(* IEC 61131-3 sources: daoli-st-library/DL_Device (part 8) *)

(* ---- FC_DL_BatteryBackupTimeCalc.st ---- *)
(*
 * FC_DL_BatteryBackupTimeCalc | C2 | DL_Device
 * 功能：电池组恒功率放电后备时间（含寿命末期与放电效率修正）       单位：容量 [Ah]、电压 [V]、功率 [kW]、时间 [min]、修正系数 [1]
 * 工况边界：恒功率简化模型（不含 Peukert 效应与温度修正，温度影响由 rDerate 吸收）；负载功率须 >0（入分母），容量、电压须 >0，两修正系数须在 (0,1]；电池组按串联单体电压和计算
 * 代数值回代：C=200 Ah、V=480 V、P=100 kW、derate=0.85、eol=0.8 → 200×480×0.85×0.8=65280 Wh；65280/100000=0.6528 h=39.17 min（spec 记 39.2 min，一致）
 * 开源溯源：clean-room 自研，未复制任何第三方代码（无外部来源）
 *)
FUNCTION FC_DL_BatteryBackupTimeCalc : BOOL
VAR_INPUT
    rCapacityAh : REAL := 200.0;     // 电池组额定容量 | battery string rated capacity [Ah]
    rStringV    : REAL := 480.0;     // 电池组标称电压 | battery string nominal voltage [V]
    rLoadKw     : REAL := 100.0;     // 放电负载功率 | discharge load power [kW]
    rDerate     : REAL := 0.85;      // 放电效率与温度综合修正 | combined discharge efficiency and temperature derating [1]
    rEolFactor  : REAL := 0.8;       // 寿命末期容量保持率 | end of life capacity retention [1]
END_VAR
VAR_OUTPUT
    rBackupMin : REAL;               // 后备时间 | backup time [min]
    rEnergyWh  : REAL;               // 可用能量 | usable energy [Wh]
    xValid     : BOOL;               // 输出有效 | outputs valid
END_VAR
VAR
    xFinC   : BOOL;                  // 容量有限性 | capacity is finite
    xFinV   : BOOL;                  // 电压有限性 | voltage is finite
    xFinP   : BOOL;                  // 功率有限性 | load power is finite
    xFinDr  : BOOL;                  // 效率修正有限性 | derating factor is finite
    xFinEol : BOOL;                  // 寿命修正有限性 | end of life factor is finite
    rPW     : REAL;                  // 负载功率（W）| load power in watts [W]
END_VAR
VAR CONSTANT
    DL_BBT_MIN_PER_HOUR : REAL := 60.0;    // 小时转分系数 | hours to minutes factor [min/h]
    DL_BBT_W_PER_KW     : REAL := 1000.0;  // 千瓦转瓦系数 | kilowatts to watts factor [W/kW]
    DL_BBT_P_MIN        : REAL := 1.0E-9;  // 负载功率下限（防零除）| load power lower bound [W]
END_VAR

// 段1｜非有限闸（R19）
xFinC := (rCapacityAh = rCapacityAh) AND ((rCapacityAh - rCapacityAh) = 0.0);
xFinV := (rStringV = rStringV) AND ((rStringV - rStringV) = 0.0);
xFinP := (rLoadKw = rLoadKw) AND ((rLoadKw - rLoadKw) = 0.0);
xFinDr := (rDerate = rDerate) AND ((rDerate - rDerate) = 0.0);
xFinEol := (rEolFactor = rEolFactor) AND ((rEolFactor - rEolFactor) = 0.0);
IF (NOT xFinC) OR (NOT xFinV) OR (NOT xFinP) OR (NOT xFinDr) OR (NOT xFinEol) THEN
    rBackupMin := 0.0;               // 安全值：后备时间 0 | safe value, zero backup time
    rEnergyWh := 0.0;
    xValid := FALSE;
    FC_DL_BatteryBackupTimeCalc := FALSE;
    RETURN;
END_IF

// 段2｜域闸：容量/电压/功率须为正，两修正系数须在 (0,1]
IF (rCapacityAh <= 0.0) OR (rStringV <= 0.0) OR (rLoadKw <= 0.0)
   OR (rDerate <= 0.0) OR (rDerate > 1.0) OR (rEolFactor <= 0.0) OR (rEolFactor > 1.0) THEN
    rBackupMin := 0.0;
    rEnergyWh := 0.0;
    xValid := FALSE;
    FC_DL_BatteryBackupTimeCalc := FALSE;
    RETURN;
END_IF

// 段3｜算法：可用能量 Wh 与后备时间 min
rEnergyWh := rCapacityAh * rStringV * rDerate * rEolFactor;
rPW := rLoadKw * DL_BBT_W_PER_KW;
IF rPW > DL_BBT_P_MIN THEN
    rBackupMin := rEnergyWh / rPW * DL_BBT_MIN_PER_HOUR;
ELSE
    rBackupMin := 0.0;               // 理论不可达（段2已排除），防御性兜底 | unreachable defence
END_IF

// 段4｜出口
xValid := TRUE;
FC_DL_BatteryBackupTimeCalc := TRUE;
END_FUNCTION

(* ---- FC_DL_BoothFilterLifeCalc.st ---- *)
(*
  Name: FC_DL_BoothFilterLifeCalc
  Category: DL_Device
  Version: 1.0.0
  Round: R89 / 2026-11-25
  开源溯源：clean-room 自研（族 涂装喷涂线，ST 开源生态实测 0 命中，无外部代码引入）
  功能：过滤棉剩余寿命：按压差累积法算寿命消耗百分比，并按当前压差增长率外推剩余运行小时。
  边界条件：① 四入参全部过非有限闸，任一非有限返回哨兵 -1；
            ② 新棉压差必须 > 0 且报废压差必须高于新棉压差（否则分母 ΔP 塌零，返回哨兵 -1）；
            ③ 已用压差 Δp − Δp_new 为除子，外推前显式判零：低于 DL_EPS 时剩余小时按满寿命处理；
            ④ 寿命百分比钳 0~100 %（量值饱和）；报警门限 90 %，超报废压差即 100 % 并报警。
  量纲自证：(ΔP − ΔP_new)/(ΔP_end − ΔP_new) 无量纲；h × 无量纲 = h。
*)
FUNCTION FC_DL_BoothFilterLifeCalc : REAL
VAR_INPUT
    fDpPa : REAL;           (* 当前滤棉压差 [Pa] Current filter pressure drop [Pa] *)
    fDpNewPa : REAL;        (* 新棉压差（洁净基线） [Pa] Clean filter pressure drop [Pa] *)
    fDpEndPa : REAL;        (* 报废压差 [Pa] End-of-life pressure drop [Pa] *)
    fRunHours : REAL;       (* 滤棉已运行小时 [h] Filter accumulated run hours [h] *)
END_VAR
VAR_OUTPUT
    fLifeUsedPct : REAL;    (* 寿命消耗百分比 [%] Life used [%] *)
    fRemainHours : REAL;    (* 剩余可用小时（外推） [h] Remaining hours, extrapolated [h] *)
    xReplaceAlarm : BOOL;   (* 更换报警（寿命 ≥ 90 %） [-] Replace alarm *)
    xValid : BOOL;          (* 计算有效性标志 [-] Calculation valid flag *)
END_VAR
VAR CONSTANT
    DL_EPS : REAL := 1.0E-9;        (* 除零判定容差 [-] Divide-by-zero tolerance *)
    DL_PCT : REAL := 100.0;         (* 百分数基准 [%] Percent base *)
    DL_ALARM_PCT : REAL := 90.0;    (* 更换报警门限 [%] Replace alarm threshold [%] *)
    DL_P_NEW_MAX : REAL := 500.0;   (* 新棉压差上限 [Pa] Clean pressure ceiling [Pa] *)
    DL_P_END_MIN : REAL := 100.0;   (* 报废压差下限 [Pa] End pressure floor [Pa] *)
    DL_P_END_MAX : REAL := 5000.0;  (* 报废压差上限 [Pa] End pressure ceiling [Pa] *)
    DL_H_MAX : REAL := 100000.0;    (* 运行小时上限 [h] Run hours ceiling [h] *)
END_VAR
VAR
    fSpanPa : REAL;     (* 全寿命压差跨度 [Pa] Full-life pressure span [Pa] *)
    fUsedPa : REAL;     (* 已消耗压差 [Pa] Consumed pressure drop [Pa] *)
    fPct : REAL;        (* 寿命消耗中间量 [%] Life used scratch [%] *)
END_VAR
(* 出口预置：四出口统一预置（R256） *)
fLifeUsedPct := 0.0; fRemainHours := 0.0; xReplaceAlarm := FALSE; xValid := FALSE;
(* 非有限闸：NaN 自反判 + Inf 差值自减判，四入参全枚举 *)
IF (fDpPa <> fDpPa) OR ((fDpPa - fDpPa) <> 0.0)
   OR (fDpNewPa <> fDpNewPa) OR ((fDpNewPa - fDpNewPa) <> 0.0)
   OR (fDpEndPa <> fDpEndPa) OR ((fDpEndPa - fDpEndPa) <> 0.0)
   OR (fRunHours <> fRunHours) OR ((fRunHours - fRunHours) <> 0.0) THEN
    FC_DL_BoothFilterLifeCalc := -1.0;      (* 哨兵 -1：入参非有限 / Sentinel -1, non-finite input *)
    RETURN;
END_IF
(* 组态域闸：压差三点与运行小时定域，报废压差须高于新棉压差 *)
IF (fDpNewPa < DL_EPS) OR (fDpNewPa > DL_P_NEW_MAX)
   OR (fDpEndPa < DL_P_END_MIN) OR (fDpEndPa > DL_P_END_MAX)
   OR ((fDpEndPa - fDpNewPa) <= DL_EPS)
   OR (fDpPa < 0.0) OR (fDpPa > (fDpEndPa * 1.5))
   OR (fRunHours < 0.0) OR (fRunHours > DL_H_MAX) THEN
    FC_DL_BoothFilterLifeCalc := -1.0;      (* 哨兵 -1：组态非法 / Sentinel -1, bad configuration *)
    RETURN;
END_IF
(* 全寿命压差跨度已过正性闸，绝无零除 *)
fSpanPa := fDpEndPa - fDpNewPa;
(* 已消耗压差：低于新棉基线按 0 处理（新棉初期压差抖动不产生负寿命） *)
fUsedPa := fDpPa - fDpNewPa;
IF fUsedPa < 0.0 THEN
    fUsedPa := 0.0;
END_IF
(* 寿命消耗百分比 *)
fPct := (fUsedPa / fSpanPa) * DL_PCT;
IF fPct > DL_PCT THEN
    fPct := DL_PCT;                         (* 量值饱和：超报废压差即 100 % / Saturation at 100 % *)
END_IF
fLifeUsedPct := fPct;
(* 剩余小时外推：h × (剩余压差/已耗压差)；已耗压差塌零时按满寿命 + 无穷处置为 0 剩余待定 *)
IF fUsedPa <= DL_EPS THEN
    fRemainHours := DL_H_MAX;               (* 近乎新棉：剩余小时按可表上限 / Effectively new filter *)
ELSE
    fRemainHours := fRunHours * ((fSpanPa - fUsedPa) / fUsedPa);
    IF fRemainHours < 0.0 THEN
        fRemainHours := 0.0;                (* 已超报废压差：剩余 0 h / Past end of life *)
    END_IF
END_IF
xReplaceAlarm := fLifeUsedPct >= DL_ALARM_PCT;
xValid := TRUE;                             (* 链路有效 / Chain valid *)
FC_DL_BoothFilterLifeCalc := fLifeUsedPct;
END_FUNCTION

(* ---- FC_DL_BrgThermalDriftRate.st ---- *)
(*
  道莅工业代码库 / Daoli Industrial ST Library
  组件: FC_DL_BrgThermalDriftRate
  分类: DL_Device
  开源溯源: 无（clean-room 工程公式自研；参考公开工艺计算公式，未复制任何受版权保护代码）
  许可证: 本项目自有 (MIT)
  功能: 轴承温升速率计算、相对环境温升与温升过快判定
*)
FUNCTION FC_DL_BrgThermalDriftRate : BOOL
VAR_INPUT
    rTempNow : REAL; // 本次轴承温度 [°C] / current bearing temperature
    rTempPrev : REAL; // 上次轴承温度 [°C] / previous bearing temperature
    rDtMin : REAL; // 采样间隔 [min] / sampling interval in minutes
    rAmbC : REAL; // 环境温度 [°C] / ambient temperature
    rAlarmRisePerMin : REAL; // 温升速率报警门槛 [°C/min] / rise rate alarm threshold
END_VAR
VAR_OUTPUT
    rRisePerMin : REAL; // 温升速率 [°C/min] / temperature rise rate
    rOverAmbC : REAL; // 相对环境温升 [°C] / temperature rise above ambient
    bValid : BOOL; // 结果有效位 [-] / result valid flag
    bFastRise : BOOL; // 温升过快标志 [-] / fast rise flag
    iErrCode : INT; // 事件码 0=正常 1=采样间隔非法 2=结果非有限 / event code
END_VAR
VAR CONSTANT
    rAbsZero : REAL := -273.15; // 绝对零度 [°C] / absolute zero in Celsius
END_VAR
VAR
    rRiseRaw : REAL; // 未校验温升速率 [°C/min] / unchecked rise rate
END_VAR

    // —— 段 0：全路径预清 —— //
    rRiseRaw := 0.0;
    rRisePerMin := 0.0;
    rOverAmbC := 0.0;
    bValid := FALSE;
    bFastRise := FALSE;
    iErrCode := 0;
    FC_DL_BrgThermalDriftRate := FALSE;
    // —— 段 1：分母闸（采样间隔必须为正） —— //
    IF rDtMin <= 0.0 THEN
        iErrCode := 1; // 采样间隔非法，速率无定义 / invalid interval, rate undefined
        RETURN;
    END_IF;
    // —— 段 2：量纲链 (°C - °C)/(min) = °C/min —— //
    rRiseRaw := (rTempNow - rTempPrev) / rDtMin; // 温升速率 [°C/min] / rise rate
    IF ABS(rRiseRaw) > 1.0E15 THEN
        iErrCode := 2; // 结果非有限，强制归零 / non-finite result, forced to zero
        RETURN;
    END_IF;
    rRisePerMin := rRiseRaw;
    // —— 段 3：相对环境温升（量纲 °C - °C = °C） —— //
    IF rTempNow <= rAbsZero THEN
        iErrCode := 2; // 温度低于绝对零度，物理不可能 / temperature below absolute zero
        RETURN;
    END_IF;
    rOverAmbC := rTempNow - rAmbC; // 相对环境温升 [°C] / rise above ambient
    // —— 段 4：温升过快判定（门槛为负时按绝对值口径比对） —— //
    IF rAlarmRisePerMin > 0.0 THEN
        bFastRise := rRisePerMin > rAlarmRisePerMin; // 常规比对 / normal comparison
    ELSE
        bFastRise := rRisePerMin > ABS(rAlarmRisePerMin); // 门槛配置异常时退化为绝对值口径 / fallback on bad threshold
    END_IF;
    bValid := TRUE;
    FC_DL_BrgThermalDriftRate := TRUE;
END_FUNCTION

(* ---- FC_DL_BushingDwellFlowCalc.st ---- *)
// FC_DL_BushingDwellFlowCalc v1.0.0
// 开源溯源：clean-room 自研（族 DL_Device，ST 生态实测 0 命中，无外部代码引入）
(*
  功能: 漏孔玻璃液质量流量（Hagen-Poiseuille 圆管层流）：r = d/2/1000，L = len/1000，
        Q = π·Δp·r⁴/(8·μ·L) [m³/s]，单孔 = Q·ρ·3.6e6 [g/h]，总流量 = 单孔·孔数/1000 [kg/h]。
  邻件/码位: 与 FC_DL_FiberDiameterFromDrawRateCalc 直接串联（本件出单孔流量）；
             16#0002_9222 = 非有限、黏度/孔径/孔长/密度非正或孔数 < 1 拒收。
*)
FUNCTION FC_DL_BushingDwellFlowCalc : REAL
VAR_INPUT
    fDeltaP    : REAL := 5000.0;    // 漏板上下压差 [Pa]，域 > 0 / Pressure differential [Pa]
    fHoleDia   : REAL := 1.6;       // 漏孔直径 [mm]，域 > 0 / Orifice diameter [mm]
    fDwellLen  : REAL := 4.0;       // 漏孔长度 [mm]，域 > 0 / Orifice length [mm]
    fViscosity : REAL := 500.0;     // 玻璃液黏度 [Pa·s]，域 > 0 / Glass viscosity [Pa s]
    iHoleCount : INT := 800;        // 漏孔数，域 >= 1 [个] / Orifice count
    fDensity   : REAL := 2500.0;    // 玻璃液密度 [kg/m³]，域 > 0 / Glass density [kg/m^3]
END_VAR
VAR_OUTPUT
    fFlowPerHole : REAL;            // 单孔质量流量 [g/h] / Mass flow per orifice [g/h]
    fFlowTotal   : REAL;            // 总质量流量 [kg/h] / Total mass flow [kg/h]
    bValid       : BOOL;            // 结果有效回执 [-] / Result validity receipt
    uErrorId     : UDINT;           // 事件码，0 = 无事件 / Event code
END_VAR
VAR
    fRadius  : REAL := 0.0;         // 漏孔半径 [m] / Orifice radius [m]
    fLenM    : REAL := 0.0;         // 漏孔长度 [m] / Orifice length [m]
    fVolFlow : REAL := 0.0;         // 单孔体积流量 [m³/s] / Volumetric flow [m^3/s]
END_VAR
// 段 0：全路径出口安全缺省 / Safe defaults on all outlets
fFlowPerHole := 0.0;                // 单孔流量缺省零 / Per-orifice default zero
fFlowTotal := 0.0;                  // 总流量缺省零 / Total flow default zero
bValid := FALSE;                    // 有效回执预清 / Validity preset clear
uErrorId := 16#0000;                // 事件码预清 / Event code preset clear
FC_DL_BushingDwellFlowCalc := 0.0;  // 返回值缺省零（镜像单孔流量）/ Return default zero
// 段 1：非有限闸（五实数入参；整数入参天然有限）/ Non-finite gate on real inputs
IF (fDeltaP <> fDeltaP) OR (fHoleDia <> fHoleDia) OR (fDwellLen <> fDwellLen)
   OR (fViscosity <> fViscosity) OR (fDensity <> fDensity)
   OR (ABS(fDeltaP) >= 3.0E38) OR (ABS(fHoleDia) >= 3.0E38) OR (ABS(fDwellLen) >= 3.0E38)
   OR (ABS(fViscosity) >= 3.0E38) OR (ABS(fDensity) >= 3.0E38) THEN
    uErrorId := 16#0002_9222;   // 入参非有限拒收 / Non-finite input reject
    RETURN;
END_IF
// 段 2：域闸（黏度/孔径/孔长/密度为正防除零 + 孔数下限，R4）/ Domain gate
IF (fViscosity <= 1.0E-6) OR (fHoleDia <= 1.0E-6) OR (fDwellLen <= 1.0E-6) OR (fDensity <= 1.0E-6) THEN
    uErrorId := 16#0002_9222;   // 黏度、孔径、孔长或密度非正 / Non-positive physical input
    RETURN;
END_IF
IF iHoleCount < 1 THEN
    uErrorId := 16#0002_9222;   // 孔数不足 1 / Orifice count below one
    RETURN;
END_IF
// 段 3：主计算（半径/长度换算 → 体积流量 → 质量流量）/ Main computation
fRadius := fHoleDia / 2.0 / 1000.0;                             // 半径 [m] / Radius in metres
fLenM := fDwellLen / 1000.0;                                    // 孔长 [m] / Length in metres
fVolFlow := 3.14159265358979 * fDeltaP * fRadius * fRadius * fRadius * fRadius
          / (8.0 * fViscosity * fLenM);                         // Q = πΔp r⁴/(8μL) / Poiseuille flow
fFlowPerHole := fVolFlow * fDensity * 3600.0 * 1000.0;          // 单孔 [g/h] / Per-orifice mass flow
fFlowTotal := fFlowPerHole * INT_TO_REAL(iHoleCount) / 1000.0;  // 总流量 [kg/h] / Total mass flow
// 段 4：出口闸（双输出非有限复核 + 非负复核）/ Outlet gate
IF (fFlowPerHole <> fFlowPerHole) OR (fFlowTotal <> fFlowTotal)
   OR (ABS(fFlowPerHole) >= 3.0E38) OR (ABS(fFlowTotal) >= 3.0E38)
   OR (fFlowPerHole < 0.0) OR (fFlowTotal < 0.0) THEN
    fFlowPerHole := 0.0;        // 复核失败回缺省 / Fallback on recheck failure
    fFlowTotal := 0.0;          // 复核失败回缺省 / Fallback on recheck failure
    uErrorId := 16#0002_9222;   // 出口复核拒收 / Output recheck reject
    RETURN;
END_IF
bValid := TRUE;                 // 有效回执 / Validity receipt
FC_DL_BushingDwellFlowCalc := fFlowPerHole;     // 返回值镜像单孔流量 / Return mirrors flow
END_FUNCTION

(* ---- FC_DL_BushingPowerBalanceCalc.st ---- *)
// FC_DL_BushingPowerBalanceCalc v1.0.0
// 开源溯源：clean-room 自研（族 DL_Device，ST 生态实测 0 命中，无外部代码引入）
(*
  功能: 漏板电热功率平衡：输入功率 = I²·R [W]→[kW]（mΩ 除 1000 转 Ω，W 除 1000 转 kW），
        对流 = 12·A·ΔT/1000 [kW]（12 为自然对流综合换热系数 W/(m²·K)），
        辐射 = εσ·A·(T_K⁴ − Ta_K⁴)/1000 [kW]（ε = 0.85，σ = 5.67e-8），
        热效率 = 1 − (对流 + 辐射)/输入功率。
  邻件/码位: 与 FC_DL_BushingTempZoneCalc 为热平衡两侧（温度设定 vs 实际电功率与散热）；
             16#0002_9227 = 非有限、电阻/面积非正、温度不高于绝对零度、输入功率近零或效率出物理域。
*)
FUNCTION FC_DL_BushingPowerBalanceCalc : REAL
VAR_INPUT
    fCurrent     : REAL := 300.0;   // 漏板电流 [A]，域 > 0 / Bushing current [A]
    fResistance  : REAL := 30.0;    // 漏板电阻 [mΩ]，域 > 0 / Bushing resistance [mOhm]
    fSurfaceArea : REAL := 0.5;     // 漏板表面积 [m²]，域 > 0 / Surface area [m^2]
    fTemp        : REAL := 1200.0;  // 漏板温度 [°C] / Bushing temperature [degC]
    fAmbient     : REAL := 30.0;    // 环境温度 [°C] / Ambient temperature [degC]
END_VAR
VAR_OUTPUT
    fPowerIn    : REAL;             // 输入电功率 [kW] / Electrical input power [kW]
    fLossConv   : REAL;             // 对流散热 [kW] / Convective loss [kW]
    fLossRad    : REAL;             // 辐射散热 [kW] / Radiative loss [kW]
    fEfficiency : REAL;             // 热效率 [-] / Thermal efficiency
    bValid      : BOOL;             // 结果有效回执 [-] / Result validity receipt
    uErrorId    : UDINT;            // 事件码，0 = 无事件 / Event code
END_VAR
VAR
    fTK  : REAL := 0.0;             // 板绝对温度 [K] / Bushing absolute temperature [K]
    fTaK : REAL := 0.0;             // 环境绝对温度 [K] / Ambient absolute temperature [K]
END_VAR
// 段 0：全路径出口安全缺省 / Safe defaults on all outlets
fPowerIn := 0.0;                    // 输入功率缺省零 / Input power default zero
fLossConv := 0.0;                   // 对流散热缺省零 / Convective loss default zero
fLossRad := 0.0;                    // 辐射散热缺省零 / Radiative loss default zero
fEfficiency := 0.0;                 // 热效率缺省零 / Efficiency default zero
bValid := FALSE;                    // 有效回执预清 / Validity preset clear
uErrorId := 16#0000;                // 事件码预清 / Event code preset clear
FC_DL_BushingPowerBalanceCalc := 0.0;   // 返回值缺省零（镜像热效率）/ Return default zero
// 段 1：非有限闸（五入参全枚举）/ Non-finite gate over all inputs
IF (fCurrent <> fCurrent) OR (fResistance <> fResistance) OR (fSurfaceArea <> fSurfaceArea)
   OR (fTemp <> fTemp) OR (fAmbient <> fAmbient)
   OR (ABS(fCurrent) >= 3.0E38) OR (ABS(fResistance) >= 3.0E38) OR (ABS(fSurfaceArea) >= 3.0E38)
   OR (ABS(fTemp) >= 3.0E38) OR (ABS(fAmbient) >= 3.0E38) THEN
    uErrorId := 16#0002_9227;   // 入参非有限拒收 / Non-finite input reject
    RETURN;
END_IF
// 段 2：域闸（电阻/面积为正 + 温度高于绝对零度 + 输入功率近零，R4）/ Domain gate
IF (fResistance <= 1.0E-6) OR (fSurfaceArea <= 1.0E-6) THEN
    uErrorId := 16#0002_9227;   // 电阻或面积非正 / Non-positive resistance or area
    RETURN;
END_IF
IF (fTemp <= -273.15) OR (fAmbient <= -273.15) THEN
    uErrorId := 16#0002_9227;   // 温度不高于绝对零度，四次方无意义 / At or below absolute zero
    RETURN;
END_IF
fPowerIn := fCurrent * fCurrent * (fResistance / 1000.0) / 1000.0;      // I²R [kW] / Input power
IF fPowerIn <= 1.0E-6 THEN
    uErrorId := 16#0002_9227;   // 输入功率近零，效率不可解 / Input power too small
    RETURN;
END_IF
// 段 3：主计算（对流 + 辐射 + 效率）/ Main computation
fTK := fTemp + 273.15;                                          // 板绝对温度 [K] / Absolute temperature
fTaK := fAmbient + 273.15;                                      // 环境绝对温度 [K] / Ambient absolute temperature
fLossConv := 12.0 * fSurfaceArea * (fTemp - fAmbient) / 1000.0;  // 对流散热 [kW] / Convective loss
fLossRad := 5.67E-8 * 0.85 * fSurfaceArea * ((fTK * fTK * fTK * fTK) - (fTaK * fTaK * fTaK * fTaK)) / 1000.0;
fEfficiency := 1.0 - (fLossConv + fLossRad) / fPowerIn;         // 热效率 / Thermal efficiency
// 段 4：出口闸（四输出非有限复核 + 效率区间复核）/ Outlet gate
IF (fPowerIn <> fPowerIn) OR (fLossConv <> fLossConv) OR (fLossRad <> fLossRad)
   OR (fEfficiency <> fEfficiency)
   OR (ABS(fPowerIn) >= 3.0E38) OR (ABS(fLossConv) >= 3.0E38)
   OR (ABS(fLossRad) >= 3.0E38) OR (ABS(fEfficiency) >= 3.0E38) THEN
    fPowerIn := 0.0;            // 复核失败回缺省 / Fallback on recheck failure
    fLossConv := 0.0;           // 复核失败回缺省 / Fallback on recheck failure
    fLossRad := 0.0;            // 复核失败回缺省 / Fallback on recheck failure
    fEfficiency := 0.0;         // 复核失败回缺省 / Fallback on recheck failure
    uErrorId := 16#0002_9227;   // 出口非有限拒收 / Output non-finite reject
    RETURN;
END_IF
IF (fEfficiency > 1.0) OR (fEfficiency < -1.0) THEN
    uErrorId := 16#0002_9227;   // 信息级：效率出物理域 / Info: efficiency out of physical range
    RETURN;                     // bValid 保持 FALSE / Validity stays false
END_IF
bValid := TRUE;                 // 有效回执 / Validity receipt
FC_DL_BushingPowerBalanceCalc := fEfficiency;   // 返回值镜像热效率 / Return mirrors efficiency
END_FUNCTION

(* ---- FC_DL_BushingTempZoneCalc.st ---- *)
// FC_DL_BushingTempZoneCalc v1.0.0
// 开源溯源：clean-room 自研（族 DL_Device，ST 生态实测 0 命中，无外部代码引入）
(*
  功能: 漏板分区温度设定：偏移 = 梯度·(iZoneIndex − (iZoneCount−1)/2)，温度 = 基准 + 偏移；
        以区号相对中心对称取偏移，保证漏板横向温度对称分布。
  邻件/码位: 与 FC_DL_BushingDwellFlowCalc（温度→黏度→流量）上游衔接；
             16#0002_9221 = 非有限、区数非正、区号越界或温度出 1100~1350 °C 拒收。
*)
FUNCTION FC_DL_BushingTempZoneCalc : REAL
VAR_INPUT
    fBaseTemp  : REAL := 1250.0;    // 中心区设定温度 [°C] / Center zone setpoint [degC]
    fGradient  : REAL := 5.0;       // 区间梯度 [°C/区] / Per-zone gradient [degC/zone]
    iZoneIndex : INT := 0;          // 区号，0 起 [-] / Zone index, zero based
    iZoneCount : INT := 1;          // 总区数，域 > 0 [-] / Total zone count
END_VAR
VAR_OUTPUT
    fZoneTemp : REAL;               // 分区温度设定 [°C] / Zone temperature setpoint [degC]
    bValid    : BOOL;               // 结果有效回执 [-] / Result validity receipt
    uErrorId  : UDINT;              // 事件码，0 = 无事件 / Event code
END_VAR
VAR
    fCenter : REAL := 0.0;          // 中心区号（可为半整数）[-] / Center zone position
END_VAR
// 段 0：全路径出口安全缺省 / Safe defaults on all outlets
fZoneTemp := 0.0;               // 分区温度缺省零 / Zone temperature default zero
bValid := FALSE;                // 有效回执预清 / Validity preset clear
uErrorId := 16#0000;            // 事件码预清 / Event code preset clear
FC_DL_BushingTempZoneCalc := 0.0;       // 返回值缺省零（镜像分区温度）/ Return default zero
// 段 1：非有限闸（两实数入参；整数入参天然有限）/ Non-finite gate on real inputs
IF (fBaseTemp <> fBaseTemp) OR (fGradient <> fGradient)
   OR (ABS(fBaseTemp) >= 3.0E38) OR (ABS(fGradient) >= 3.0E38) THEN
    uErrorId := 16#0002_9221;   // 入参非有限拒收 / Non-finite input reject
    RETURN;
END_IF
// 段 2：域闸（区数为正 + 区号不越界）/ Domain gate
IF iZoneCount <= 0 THEN
    uErrorId := 16#0002_9221;   // 区数非正 / Non-positive zone count
    RETURN;
END_IF
IF (iZoneIndex < 0) OR (iZoneIndex >= iZoneCount) THEN
    uErrorId := 16#0002_9221;   // 区号越界 / Zone index out of range
    RETURN;
END_IF
// 段 3：主计算（中心对称偏移）/ Main computation
fCenter := INT_TO_REAL(iZoneCount - 1) / 2.0;                   // 中心区号 / Center zone position
fZoneTemp := fBaseTemp + fGradient * (INT_TO_REAL(iZoneIndex) - fCenter);   // 分区温度 / Zone temperature
// 段 4：出口闸（非有限复核 + 1100~1350 °C 工艺窗判定）/ Outlet gate
IF (fZoneTemp <> fZoneTemp) OR (ABS(fZoneTemp) >= 3.0E38) THEN
    fZoneTemp := 0.0;           // 复核失败回缺省 / Fallback on recheck failure
    uErrorId := 16#0002_9221;   // 出口非有限拒收 / Output non-finite reject
    RETURN;
END_IF
IF (fZoneTemp < 1100.0) OR (fZoneTemp > 1350.0) THEN
    uErrorId := 16#0002_9221;   // 信息级：温度出工艺窗 / Info: temperature out of window
    RETURN;                     // bValid 保持 FALSE / Validity stays false
END_IF
bValid := TRUE;                 // 有效回执 / Validity receipt
FC_DL_BushingTempZoneCalc := fZoneTemp;     // 返回值镜像分区温度 / Return mirrors temperature
END_FUNCTION

(* ---- FC_DL_CakeMoistureDryCalc.st ---- *)
// FC_DL_CakeMoistureDryCalc v1.0.0
// 开源溯源：clean-room 自研（族 DL_Device，ST 生态实测 0 命中，无外部代码引入）
(*
  功能: 丝饼含水率与干燥时长：当前含水率 = 100·(湿重 − 干重)/湿重 [%]，
        当前水质量 = 湿重 − 干重，目标水质量 = 干重·目标/(100 − 目标)（目标按湿基反解），
        待除水 = 当前水 − 目标水（负值归零），预计时长 = 待除水/干燥速率 [h]。
  邻件/码位: 与 FC_DL_FiberCoolingAirflowCalc 同属后处理热工件（成品干燥 vs 在线冷却）；
             16#0002_9229 = 非有限、湿重不大于干重、目标含水率越界或速率非正拒收。
*)
FUNCTION FC_DL_CakeMoistureDryCalc : REAL
VAR_INPUT
    fWetMass        : REAL := 20.0;     // 湿饼质量 [kg]，域 > 干重 / Wet cake mass [kg]
    fDryMass        : REAL := 14.0;     // 干基质量 [kg]，域 >= 0 / Dry basis mass [kg]
    fTargetMoisture : REAL := 8.0;      // 目标含水率 [%]，域 [0, 100) / Target moisture [%]
    fDryRate        : REAL := 3.0;      // 干燥速率 [kg/h]，域 > 0 / Drying rate [kg/h]
END_VAR
VAR_OUTPUT
    fMoistureNow   : REAL;              // 当前含水率 [%] / Current moisture [%]
    fWaterToRemove : REAL;              // 待除水质量 [kg] / Water to remove [kg]
    fDryTimeH      : REAL;              // 预计干燥时长 [h] / Estimated drying time [h]
    bValid         : BOOL;              // 结果有效回执 [-] / Result validity receipt
    uErrorId       : UDINT;             // 事件码，0 = 无事件 / Event code
END_VAR
VAR
    fWaterNow    : REAL := 0.0;         // 当前水质量 [kg] / Current water mass [kg]
    fWaterTarget : REAL := 0.0;         // 目标水质量 [kg] / Target water mass [kg]
END_VAR
// 段 0：全路径出口安全缺省 / Safe defaults on all outlets
fMoistureNow := 0.0;                // 含水率缺省零 / Moisture default zero
fWaterToRemove := 0.0;              // 待除水缺省零 / Water to remove default zero
fDryTimeH := 0.0;                   // 干燥时长缺省零 / Drying time default zero
bValid := FALSE;                    // 有效回执预清 / Validity preset clear
uErrorId := 16#0000;                // 事件码预清 / Event code preset clear
FC_DL_CakeMoistureDryCalc := 0.0;   // 返回值缺省零（镜像待除水）/ Return default zero
// 段 1：非有限闸（四入参全枚举）/ Non-finite gate over all inputs
IF (fWetMass <> fWetMass) OR (fDryMass <> fDryMass)
   OR (fTargetMoisture <> fTargetMoisture) OR (fDryRate <> fDryRate)
   OR (ABS(fWetMass) >= 3.0E38) OR (ABS(fDryMass) >= 3.0E38)
   OR (ABS(fTargetMoisture) >= 3.0E38) OR (ABS(fDryRate) >= 3.0E38) THEN
    uErrorId := 16#0002_9229;   // 入参非有限拒收 / Non-finite input reject
    RETURN;
END_IF
// 段 2：域闸（湿重大于干重且为正 + 干基非负 + 目标区间 + 速率正，R4）/ Domain gate
IF (fWetMass <= 1.0E-6) OR (fWetMass <= fDryMass) THEN
    uErrorId := 16#0002_9229;   // 湿重非正或不大于干重 / Wet mass not above dry mass
    RETURN;
END_IF
IF fDryMass < 0.0 THEN
    uErrorId := 16#0002_9229;   // 干基质量为负 / Negative dry mass
    RETURN;
END_IF
IF (fTargetMoisture < 0.0) OR (fTargetMoisture >= 100.0) THEN
    uErrorId := 16#0002_9229;   // 目标含水率越界（分母近零）/ Target moisture out of range
    RETURN;
END_IF
IF fDryRate <= 1.0E-6 THEN
    uErrorId := 16#0002_9229;   // 干燥速率非正 / Non-positive drying rate
    RETURN;
END_IF
// 段 3：主计算（当前含水率 → 目标水 → 待除水 → 时长）/ Main computation
fWaterNow := fWetMass - fDryMass;                               // 当前水质量 [kg] / Current water
fMoistureNow := 100.0 * fWaterNow / fWetMass;                   // 当前含水率 [%] / Current moisture
fWaterTarget := fDryMass * fTargetMoisture / (100.0 - fTargetMoisture);     // 目标水 [kg] / Target water
fWaterToRemove := fWaterNow - fWaterTarget;                     // 待除水 [kg] / Water to remove
IF fWaterToRemove < 0.0 THEN
    fWaterToRemove := 0.0;                                      // 已达标归零 / Already dry, clamp zero
END_IF
fDryTimeH := fWaterToRemove / fDryRate;                         // 预计时长 [h] / Estimated time
// 段 4：出口闸（三输出非有限复核 + 非负复核）/ Outlet gate
IF (fMoistureNow <> fMoistureNow) OR (fWaterToRemove <> fWaterToRemove) OR (fDryTimeH <> fDryTimeH)
   OR (ABS(fMoistureNow) >= 3.0E38) OR (ABS(fWaterToRemove) >= 3.0E38) OR (ABS(fDryTimeH) >= 3.0E38)
   OR (fMoistureNow < 0.0) OR (fWaterToRemove < 0.0) OR (fDryTimeH < 0.0) THEN
    fMoistureNow := 0.0;        // 复核失败回缺省 / Fallback on recheck failure
    fWaterToRemove := 0.0;      // 复核失败回缺省 / Fallback on recheck failure
    fDryTimeH := 0.0;           // 复核失败回缺省 / Fallback on recheck failure
    uErrorId := 16#0002_9229;   // 出口复核拒收 / Output recheck reject
    RETURN;
END_IF
bValid := TRUE;                 // 有效回执 / Validity receipt
FC_DL_CakeMoistureDryCalc := fWaterToRemove;    // 返回值镜像待除水 / Return mirrors water
END_FUNCTION

(* ---- FC_DL_CementMillLoadCalc.st ---- *)
(*
  DL Factory R84 | FC_DL_CementMillLoadCalc
  功能：算管磨机填充率与循环负荷，并按目标区间判合格
  开源溯源：无（clean-room 自研，依据公开工艺公式，来源=行业通用公式，许可证=MIT，借鉴点=公式结构）
  规则：R1-R16 全遵守
*)
FUNCTION FC_DL_CementMillLoadCalc : REAL
VAR_INPUT
    fBallChargeT : REAL := 120.0; // 磨内钢球装载量 [t] / grinding ball charge mass [t]
    fMillVolM3 : REAL := 100.0; // 磨机有效容积 [m³] / effective mill volume [m^3]
    fBulkDensityTm3 : REAL := 4.6; // 钢球堆密度 [t/m³] / ball bulk density [t/m^3]
    fRejectTph : REAL := 120.0; // 选粉机返料（粗粉）量 [t/h] / separator rejects [t/h]
    fProductTph : REAL := 100.0; // 成品产量 [t/h] / finished product rate [t/h]
    fFillLoPct : REAL := 24.0; // 填充率合格下限 [%] / filling degree lower bound [%]
    fFillHiPct : REAL := 32.0; // 填充率合格上限 [%] / filling degree upper bound [%]
END_VAR
VAR_OUTPUT
    fCircLoad : REAL; // 循环负荷（返料/成品） [-] / circulating load ratio [-]
    xPass : BOOL; // 填充率落在目标区间 [-] / filling degree inside the band [-]
    xValid : BOOL; // 计算结果有效标志 [-] / calculation valid flag [-]
END_VAR
VAR
    fFillPct : REAL; // 填充率中间量 [%] / filling degree intermediate [%]
    fBallVolM3 : REAL; // 钢球堆积体积 [m³] / ball bulk volume [m^3]
END_VAR

// 段 1｜出口预置（R256）
FC_DL_CementMillLoadCalc := -1.0; // 哨兵返回 -1（无效） [-] / sentinel return -1, invalid [-]
fCircLoad := 0.0; // 循环负荷预置零 [-] / circulating load preset zero [-]
xPass := FALSE; // 合格位预置 FALSE [-] / pass preset false [-]
xValid := FALSE; // 计算完成前不认结果 [-] / unusable before calculation [-]

// 段 2｜非有限拦截 + 域闸（R4/R20）
IF NOT (fBallChargeT > -1.0E30 AND fBallChargeT < 1.0E30) OR NOT (fMillVolM3 > -1.0E30 AND fMillVolM3 < 1.0E30) OR NOT (fBulkDensityTm3 > -1.0E30 AND fBulkDensityTm3 < 1.0E30) THEN
    RETURN; // 装载量/容积/堆密度任一非有限即拒算 [-] / any non finite charge, volume or density rejected [-]
END_IF
IF NOT (fRejectTph > -1.0E30 AND fRejectTph < 1.0E30) OR NOT (fProductTph > -1.0E30 AND fProductTph < 1.0E30) OR NOT (fFillLoPct > -1.0E30 AND fFillLoPct < 1.0E30) OR NOT (fFillHiPct > -1.0E30 AND fFillHiPct < 1.0E30) THEN
    RETURN; // 返料/成品/区间任一非有限即拒算 [-] / any non finite flow or band rejected [-]
END_IF
IF fMillVolM3 < 1.0E-9 OR fBulkDensityTm3 < 1.0E-9 OR fProductTph < 1.0E-9 OR fBallChargeT < 0.0 OR fRejectTph < 0.0 THEN
    RETURN; // 容积/堆密度/产量正域分母闸（防除零） [m³, t/m³, t/h] / positive denominator gate [-]
END_IF
IF NOT (fFillLoPct < fFillHiPct) THEN
    RETURN; // 目标区间组态闸：下限必须严格小于上限 [%] / band config gate [%]
END_IF

// 段 3｜填充率 = 装载量 / (容积 × 钢球堆密度)
fBallVolM3 := fBallChargeT / fBulkDensityTm3; // t ÷ t/m³ = m³ / [t] / [t/m^3] = [m^3]
fFillPct := (fBallVolM3 / fMillVolM3) * 100.0; // m³ ÷ m³ × 100 = % / [m^3] / [m^3] × 100 = [%]
IF NOT (fFillPct > -1.0E30 AND fFillPct < 1.0E30) THEN
    RETURN; // 结果非有限再拦一次 [-] / second finiteness gate [-]
END_IF

// 段 4｜循环负荷 = 返料 / 成品，与区间判定
fCircLoad := fRejectTph / fProductTph; // t/h ÷ t/h = 无量纲 / [t/h] / [t/h] = [-]
IF NOT (fCircLoad > -1.0E30 AND fCircLoad < 1.0E30) THEN
    RETURN; // 结果非有限再拦一次 [-] / second finiteness gate [-]
END_IF
xPass := (fFillPct >= fFillLoPct) AND (fFillPct <= fFillHiPct); // 双边直比，禁浮点等值 [-] / two sided band compare [-]
xValid := TRUE; // 链路有效 [-] / chain valid [-]
FC_DL_CementMillLoadCalc := fFillPct; // 返回填充率 [%] / return the filling degree [%]
END_FUNCTION

(* ---- FC_DL_ChilledWaterDeltaTCalc.st ---- *)
(*
 * FC_DL_ChilledWaterDeltaTCalc | C1 | DL_Device
 * 功能：冷冻水供回水温差与「目标温差下的需求流量」互算       单位：冷量 [kW]、流量 [m³/h]、密度 [kg/m³]、比热 [kJ/(kg·K)]、温差 [K]
 * 工况边界：热平衡式 Q=ρ·cp·V̇·ΔT，cp 取 4.186 kJ/(kg·K)、ρ 取 1000 kg/m³（纯水 20 ℃）；流量须 >0 且有限；含乙二醇或高温水须重标 ρ/cp
 * 代数值回代：Q=100 kW、V=17.2 m³/h → V̇=0.004778 m³/s → ΔT=100/(1000×0.004778×4.186)=5.00 K；反算目标 5 K 时流量 17.2 m³/h（闭环自洽，与 spec 回代值 5.0 K 一致）
 * 量纲修正说明：spec 原式写作 100000/(ρ·cp·V̇) 并以 kJ 级 cp=4.186 代入，分子分母相差 1000 倍；本件按 spec 回代值 ΔT=5.0 K 采用 kW 与 kJ 同阶一致式（分子取 kW，不乘 1000）
 * 开源溯源：clean-room 自研，未复制任何第三方代码（无外部来源）
 *)
FUNCTION FC_DL_ChilledWaterDeltaTCalc : BOOL
VAR_INPUT
    rLoadKw         : REAL := 100.0;   // 冷冻水侧冷负荷 | chilled water cooling load [kW]
    rFlowM3h        : REAL := 17.2;    // 冷冻水体积流量 | chilled water volume flow [m³/h]
    rRho            : REAL := 1000.0;  // 水密度 | water density [kg/m³]
    rCp             : REAL := 4.186;   // 水定压比热 | water specific heat [kJ/(kg·K)]
    rTargetDeltaTK  : REAL := 5.0;     // 目标温差（用于反算需求流量；spec 未列，按 5 K 缺省）| target delta T for the flow back-calculation [K]
END_VAR
VAR_OUTPUT
    rDeltaTK          : REAL;          // 实际供回水温差 | actual supply to return temperature difference [K]
    rFlowForTargetM3h : REAL;          // 目标温差下的需求流量 | flow required for the target delta T [m³/h]
    xValid            : BOOL;          // 输出有效 | outputs valid
END_VAR
VAR
    xFinQ  : BOOL;                     // 冷负荷有限性 | load is finite
    xFinV  : BOOL;                     // 流量有限性 | flow is finite
    xFinR  : BOOL;                     // 密度有限性 | density is finite
    xFinCp : BOOL;                     // 比热有限性 | specific heat is finite
    xFinTg : BOOL;                     // 目标温差有限性 | target delta T is finite
    rVolM3s : REAL;                    // 体积流量（m³/s）| volume flow in SI units [m³/s]
    rCapKwPerK : REAL;                 // 热容流率 ρ×cp×V̇ | thermal capacity flow rate [kW/K]
END_VAR
VAR CONSTANT
    DL_CWD_SEC_PER_HOUR : REAL := 3600.0;  // 小时转秒系数 | hours to seconds factor [s/h]
    DL_CWD_CAP_MIN      : REAL := 1.0E-9;  // 除零保护阈值 | division guard threshold [kW/K]
END_VAR

// 段1｜非有限闸（R19）
xFinQ := (rLoadKw = rLoadKw) AND ((rLoadKw - rLoadKw) = 0.0);
xFinV := (rFlowM3h = rFlowM3h) AND ((rFlowM3h - rFlowM3h) = 0.0);
xFinR := (rRho = rRho) AND ((rRho - rRho) = 0.0);
xFinCp := (rCp = rCp) AND ((rCp - rCp) = 0.0);
xFinTg := (rTargetDeltaTK = rTargetDeltaTK) AND ((rTargetDeltaTK - rTargetDeltaTK) = 0.0);
IF (NOT xFinQ) OR (NOT xFinV) OR (NOT xFinR) OR (NOT xFinCp) OR (NOT xFinTg) THEN
    rDeltaTK := 0.0;                 // 安全值：温差 0 | safe value, zero delta T
    rFlowForTargetM3h := 0.0;
    xValid := FALSE;
    FC_DL_ChilledWaterDeltaTCalc := FALSE;
    RETURN;
END_IF

// 段2｜域闸：流量/密度/比热/目标温差均须为正（全部入分母链）
IF (rFlowM3h <= 0.0) OR (rRho <= 0.0) OR (rCp <= 0.0) OR (rTargetDeltaTK <= 0.0)
   OR (rLoadKw < 0.0) THEN
    rDeltaTK := 0.0;
    rFlowForTargetM3h := 0.0;
    xValid := FALSE;
    FC_DL_ChilledWaterDeltaTCalc := FALSE;
    RETURN;
END_IF

// 段3｜实际温差：ΔT = Q/(ρ×cp×V̇)，V̇ 由 m³/h 换算为 m³/s
rVolM3s := rFlowM3h / DL_CWD_SEC_PER_HOUR;
rCapKwPerK := rRho * rCp * rVolM3s;
IF rCapKwPerK > DL_CWD_CAP_MIN THEN
    rDeltaTK := rLoadKw / rCapKwPerK;
ELSE
    rDeltaTK := 0.0;                 // 理论不可达（段2已排除），防御性兜底 | unreachable defence
END_IF

// 段4｜反算目标温差下的需求流量：V = 3600×Q/(ρ×cp×ΔT_target)
rFlowForTargetM3h := DL_CWD_SEC_PER_HOUR * rLoadKw / (rRho * rCp * rTargetDeltaTK);
xValid := TRUE;
FC_DL_ChilledWaterDeltaTCalc := TRUE;
END_FUNCTION

(* ---- FC_DL_ChipLoadPerToothCalc.st ---- *)
(*
  DL Factory R84 | FC_DL_ChipLoadPerToothCalc
  功能：算每齿进给 fz 与切屑厚度 hm，并判最小切屑厚度以下的风险位
  开源溯源：无（clean-room 自研，依据公开工艺公式，来源=行业通用公式，许可证=MIT，借鉴点=公式结构）
  规则：R1-R16 全遵守
*)
FUNCTION FC_DL_ChipLoadPerToothCalc : REAL
VAR_INPUT
    fVf : REAL := 800.0; // 进给速度 [mm/min] / feed rate [mm/min]
    iTeeth : INT := 4; // 刀齿数（≥1） [齿] / tooth count [teeth]
    fRpm : REAL := 6000.0; // 主轴转速 [r/min] / spindle speed [r/min]
    fKrDeg : REAL := 60.0; // 主偏角 [°] / entering angle [deg]
    fMinChipMm : REAL := 0.02; // 最小切屑厚度（颤振/摩擦判据） [mm] / minimum chip thickness [mm]
END_VAR
VAR_OUTPUT
    fChipThkMm : REAL; // 切屑厚度 hm [mm] / chip thickness [mm]
    xThinChip : BOOL; // 切屑过薄风险位（摩擦/加工硬化） [-] / thin chip risk flag [-]
    xValid : BOOL; // 计算结果有效标志 [-] / calculation valid flag [-]
END_VAR
VAR
    fTeeth : REAL; // 齿数实数化 [齿] / tooth count as a real [teeth]
    fFzRaw : REAL; // 每齿进给中间量 [mm/z] / feed per tooth intermediate [mm/z]
    fKrRad : REAL; // 主偏角弧度值 [rad] / entering angle in radians [rad]
END_VAR
VAR CONSTANT
    DL_CHIP_DEG2RAD : REAL := 0.0174532925199433; // 度转弧度常量 [rad/°] / degree to radian constant [rad/deg]
END_VAR

// 段 1｜出口预置（R256）
FC_DL_ChipLoadPerToothCalc := -1.0; // 哨兵返回 -1（无效） [-] / sentinel return -1, invalid [-]
fChipThkMm := 0.0; // 切屑厚度预置零 [mm] / chip thickness preset zero [mm]
xThinChip := FALSE; // 过薄风险位预置 FALSE [-] / thin chip flag preset false [-]
xValid := FALSE; // 计算完成前不认结果 [-] / unusable before calculation [-]

// 段 2｜非有限拦截 + 域闸（R4/R20）
IF NOT (fVf > -1.0E30 AND fVf < 1.0E30) OR NOT (fRpm > -1.0E30 AND fRpm < 1.0E30) OR NOT (fKrDeg > -1.0E30 AND fKrDeg < 1.0E30) OR NOT (fMinChipMm > -1.0E30 AND fMinChipMm < 1.0E30) THEN
    RETURN; // 任一入参为 NaN/Inf 一律拒绝 [-] / any NaN or Inf input rejected [-]
END_IF
IF iTeeth < 1 OR iTeeth > 200 OR fVf < 0.0 OR fRpm < 1.0E-9 THEN
    RETURN; // 齿数与转速正域闸（防除零） [齿, r/min] / tooth count and speed gate [teeth, r/min]
END_IF
IF fKrDeg <= 0.0 OR fKrDeg >= 180.0 THEN
    RETURN; // 主偏角开区间域闸 [°] / entering angle open interval gate [deg]
END_IF

// 段 3｜fz = vf / (z × n)
fTeeth := INT_TO_REAL(iTeeth); // 标准转换，禁构造函数式 [齿] / standard conversion only [teeth]
fFzRaw := fVf / (fTeeth * fRpm); // mm/min ÷ (齿 × r/min) = mm/z / [mm/min] / ([teeth] × [r/min]) = [mm/tooth]
IF fFzRaw < 0.0 OR NOT (fFzRaw > -1.0E30 AND fFzRaw < 1.0E30) THEN
    RETURN; // 结果非有限或负值即非法 [mm/z] / non finite or negative result [mm/z]
END_IF

// 段 4｜hm = fz × sin(Kr)
fKrRad := fKrDeg * DL_CHIP_DEG2RAD; // ° × rad/° = rad / [deg] × [rad/deg] = [rad]
fChipThkMm := fFzRaw * SIN(fKrRad); // mm/z × 无量纲 = mm / [mm/tooth] × [-] = [mm]
IF NOT (fChipThkMm > -1.0E30 AND fChipThkMm < 1.0E30) THEN
    RETURN; // 结果非有限再拦一次 [-] / second finiteness gate [-]
END_IF
xThinChip := fChipThkMm < fMinChipMm; // 直比下限，禁浮点等值 [-] / direct compare against the floor [-]
xValid := TRUE; // 链路有效 [-] / chain valid [-]
FC_DL_ChipLoadPerToothCalc := fFzRaw; // 返回每齿进给 [mm/z] / return the feed per tooth [mm/tooth]
END_FUNCTION

(* ---- FC_DL_ChlorineDpdAbsorbCalc.st ---- *)
(* ============================================================
   DL_Device / FC_DL_ChlorineDpdAbsorbCalc ｜ v1.0.0 ｜ 2026-11-25
   功能：DPD 比色吸光度 → 余氯。slope = 满量程浓度 / 满量程吸光度 [mg/L per AU]，
         C = slope · (A_meas − A_zero)，再按量程钳制。
   边界：满量程吸光度 ≤ 1E-6（未标定/空皿）→ 浓度与斜率同拍写 0、返回 FALSE（N1）；
         任一浮点入参非有限 → 两出口写 0、返回 FALSE；
         nRangeSel：0=低量程 2.00 mg/L、1=高量程 5.00 mg/L，其余按低量程处理并
         返回 FALSE（档位非法）。C 越出 [0, 满量程] → 钳端点并置 bOutOfRange。
         签名无出口码，闸序即归因序（非有限 → 满量程非法 → 档位非法）。
         量纲清单（N5）：吸光度 AU 无量纲；1 AU 满量程对应档位浓度；DPD 摩尔
         吸光系数已并入斜率，不再单独换算。
   依赖：仅 IEC 61131-3（无外部依赖，纯算术） ｜ 溯源：DLF-D-WATERANA
   验收：A=0.40/A_zero=0.02/A_span=1.00/档位 0 → slope=2.0、C=0.76 mg/L；
         档位 1 → slope=5.0、C=1.90 mg/L；A_span=0 → 两出口 0、返回 FALSE。
   ============================================================ *)
FUNCTION FC_DL_ChlorineDpdAbsorbCalc : BOOL
VAR_INPUT
    fAbsMeas  : REAL;  // 样品吸光度 [AU] / Absorbance of the sample
    fAbsZero  : REAL;  // 空白（零点）吸光度 [AU] / Absorbance of the blank reference
    fAbsSpan  : REAL;  // 满量程吸光度，有效域 > 1E-6 [AU] / Full scale absorbance
    nRangeSel : INT;   // 量程档位 0=2.00 mg/L 1=5.00 mg/L [-] / Measurement range selector
END_VAR
VAR_OUTPUT
    fChlorineMgL : REAL;  // 余氯浓度 [mg/L] / Free chlorine concentration
    fSlopeMgLAu  : REAL;  // 换算斜率 [mg/L per AU] / Conversion slope in mg per liter per absorbance unit
    bOutOfRange  : BOOL;  // 换算值被钳到量程端点 [-] / Value clamped to a range end
END_VAR
VAR
    _fFull : REAL;  // 档位满量程浓度 [mg/L] / Full scale concentration of the selected range
    _fSlo  : REAL;  // 斜率中间值 [mg/L per AU] / Intermediate slope value
    _fC    : REAL;  // 浓度中间值 [mg/L] / Intermediate concentration value
    _bRng  : BOOL;  // 档位非法标志 [-] / Illegal range selector flag
END_VAR
VAR CONSTANT
    DL_DPD_RANGE_LO : REAL := 2.00;    // 低量程满量程 [mg/L] / Low range full scale
    DL_DPD_RANGE_HI : REAL := 5.00;    // 高量程满量程 [mg/L] / High range full scale
    DL_DPD_EPS      : REAL := 1.0E-6;  // 满量程吸光度判零下限 [AU] / Zero floor of the full scale absorbance
END_VAR

(* 段 0：出口预置安全侧（两出口 0、越限置位，N1/N3） *)
FC_DL_ChlorineDpdAbsorbCalc := FALSE;
fChlorineMgL := 0.0;  fSlopeMgLAu := 0.0;  bOutOfRange := TRUE;
_bRng := FALSE;

(* 段 1：非有限闸（三个浮点入参；NaN 自反 + Inf 差值自减双判，R79/R272） *)
IF (fAbsMeas <> fAbsMeas) OR (fAbsZero <> fAbsZero) OR (fAbsSpan <> fAbsSpan) THEN RETURN; END_IF
(* Inf 双判须覆盖 fAbsSpan：满量程 +Inf 使斜率算成 0、浓度算成 0 却返回 TRUE（假安全） *)
IF ((fAbsMeas - fAbsMeas) <> (fAbsMeas - fAbsMeas))
   OR ((fAbsZero - fAbsZero) <> (fAbsZero - fAbsZero))
   OR ((fAbsSpan - fAbsSpan) <> (fAbsSpan - fAbsSpan)) THEN RETURN; END_IF

(* 段 2：满量程域闸（防除零，除子在段 4 才使用） *)
IF ABS(fAbsSpan) <= DL_DPD_EPS THEN RETURN; END_IF

(* 段 3：档位分派（非法按低量程，归因独立） *)
CASE nRangeSel OF
0:      _fFull := DL_DPD_RANGE_LO;
1:      _fFull := DL_DPD_RANGE_HI;
ELSE
    _fFull := DL_DPD_RANGE_LO;  _bRng := TRUE;
END_CASE

(* 段 4：斜率与浓度（除子已证 > 1E-6） *)
_fSlo := _fFull / fAbsSpan;
_fC   := _fSlo * (fAbsMeas - fAbsZero);

(* 段 5：结果复检（非有限保持段 0 安全侧） *)
IF (_fC <> _fC) OR ((_fC - _fC) <> (_fC - _fC)) THEN RETURN; END_IF

(* 段 6：单一出口裁决（判据与出口同源于 _fC 与 _fFull，N4/R23） *)
fSlopeMgLAu := _fSlo;
bOutOfRange := ((_fC < 0.0) OR (_fC > _fFull));
IF _fC < 0.0 THEN
    fChlorineMgL := 0.0;                // 负值保护：钳零后上报
ELSIF _fC > _fFull THEN
    fChlorineMgL := _fFull;             // 饱和上报：钳顶后值仍可读
ELSE
    fChlorineMgL := _fC;
END_IF
FC_DL_ChlorineDpdAbsorbCalc := NOT _bRng;    // 档位非法：值照给、返回 FALSE
END_FUNCTION

(* ---- FC_DL_ClinkerC3sCalc.st ---- *)
(*
  DL Factory R84 | FC_DL_ClinkerC3sCalc
  功能：Bogue 法算熟料 C3S 含量并附 C2S / C3A / C4AF，负值按 0 钳位
  开源溯源：无（clean-room 自研，依据公开工艺公式，来源=行业通用公式，许可证=MIT，借鉴点=公式结构）
  规则：R1-R16 全遵守
*)
FUNCTION FC_DL_ClinkerC3sCalc : REAL
VAR_INPUT
    fCaO : REAL := 65.0; // 氧化钙含量 [%] / calcium oxide content [%]
    fSiO2 : REAL := 21.0; // 二氧化硅含量 [%] / silica content [%]
    fAl2O3 : REAL := 5.2; // 三氧化二铝含量 [%] / alumina content [%]
    fFe2O3 : REAL := 3.4; // 三氧化二铁含量 [%] / ferric oxide content [%]
    fSO3 : REAL := 1.0; // 三氧化硫含量 [%] / sulfur trioxide content [%]
END_VAR
VAR_OUTPUT
    fC2s : REAL; // 硅酸二钙 C2S 含量 [%] / dicalcium silicate content [%]
    fC3a : REAL; // 铝酸三钙 C3A 含量 [%] / tricalcium aluminate content [%]
    fC4af : REAL; // 铁铝酸四钙 C4AF 含量 [%] / tetracalcium aluminoferrite content [%]
    xValid : BOOL; // 计算结果有效标志 [-] / calculation valid flag [-]
END_VAR
VAR
    fC3sRaw : REAL; // 未钳位 C3S 计算值 [%] / unclamped C3S value [%]
    fC3sClamp : REAL; // 钳位后 C3S [%] / clamped C3S [%]
    fC2sRaw : REAL; // 未钳位 C2S 计算值 [%] / unclamped C2S value [%]
    fC3aRaw : REAL; // 未钳位 C3A 计算值 [%] / unclamped C3A value [%]
    fC4afRaw : REAL; // 未钳位 C4AF 计算值 [%] / unclamped C4AF value [%]
    i : INT; // 钳位循环游标 [-] / clamp loop cursor [-]
    fArr : ARRAY[0..2] OF REAL; // 待钳位三相暂存（C2S/C3A/C4AF） [%] / staged phases for clamping [%]
END_VAR

// 段 1｜出口预置（R256）
FC_DL_ClinkerC3sCalc := -1.0; // 哨兵返回 -1（无效） [-] / sentinel return -1, invalid [-]
fC2s := 0.0; // C2S 预置零 [%] / C2S preset zero [%]
fC3a := 0.0; // C3A 预置零 [%] / C3A preset zero [%]
fC4af := 0.0; // C4AF 预置零 [%] / C4AF preset zero [%]
xValid := FALSE; // 计算完成前不认结果 [-] / unusable before calculation [-]

// 段 2｜非有限拦截 + 域闸（R4/R20）
IF NOT (fCaO > -1.0E30 AND fCaO < 1.0E30) OR NOT (fSiO2 > -1.0E30 AND fSiO2 < 1.0E30) OR NOT (fAl2O3 > -1.0E30 AND fAl2O3 < 1.0E30) OR NOT (fFe2O3 > -1.0E30 AND fFe2O3 < 1.0E30) OR NOT (fSO3 > -1.0E30 AND fSO3 < 1.0E30) THEN
    RETURN; // 五项氧化物任一非有限即拒算 [-] / any non finite oxide rejected [-]
END_IF
IF fCaO < 0.0 OR fSiO2 < 0.0 OR fAl2O3 < 0.0 OR fFe2O3 < 0.0 OR fSO3 < 0.0 THEN
    RETURN; // 化学分析值非负域闸（负含量物理非法） [%] / non negative chemical analysis gate [%]
END_IF

// 段 3｜C3S = 4.071CaO − 7.6SiO2 − 6.718Al2O3 − 1.43Fe2O3 − 2.852SO3
fC3sRaw := ((((4.071 * fCaO) - (7.6 * fSiO2)) - (6.718 * fAl2O3)) - (1.43 * fFe2O3)) - (2.852 * fSO3); // % 各项线性组合 = %（系数无量纲） / linear combination of [%] terms = [%]
IF NOT (fC3sRaw > -1.0E30 AND fC3sRaw < 1.0E30) THEN
    RETURN; // 结果非有限再拦一次 [-] / second finiteness gate [-]
END_IF

// 段 4｜C2S = 2.867SiO2 − 0.7544C3S（按未钳位 C3S 计，符合 Bogue 原式）
fC2sRaw := (2.867 * fSiO2) - (0.7544 * fC3sRaw); // % − % = % / [%] minus [%] = [%]
fC3aRaw := (2.65 * fAl2O3) - (1.692 * fFe2O3); // % − % = % / [%] minus [%] = [%]
fC4afRaw := 3.043 * fFe2O3; // % × 无量纲 = % / [%] × [-] = [%]

// 段 5｜负值钳位：四相统一走定长数组，正向游标 0→2（禁反向递减循环）
fC3sClamp := fC3sRaw; // 先接未钳位值 [%] / take the raw C3S [%]
IF fC3sClamp < 0.0 THEN
    fC3sClamp := 0.0; // C3S 负值钳零 [%] / clamp negative C3S to zero [%]
END_IF
fArr[0] := fC2sRaw; // 装入 C2S [%] / load C2S [%]
fArr[1] := fC3aRaw; // 装入 C3A [%] / load C3A [%]
fArr[2] := fC4afRaw; // 装入 C4AF [%] / load C4AF [%]
FOR i := 0 TO 2 DO
    IF fArr[i] < 0.0 THEN
        fArr[i] := 0.0; // 负值钳零（矿物含量物理非负） [%] / clamp to zero, mineral content is non negative [%]
    END_IF
END_FOR
fC2s := fArr[0]; // C2S 落定 [%] / land C2S [%]
fC3a := fArr[1]; // C3A 落定 [%] / land C3A [%]
fC4af := fArr[2]; // C4AF 落定 [%] / land C4AF [%]
xValid := TRUE; // 链路有效 [-] / chain valid [-]
FC_DL_ClinkerC3sCalc := fC3sClamp; // 返回钳位后 C3S [%] / return the clamped C3S [%]
END_FUNCTION

(* ---- FC_DL_ClinkerFreeLimeCalc.st ---- *)
(*
  DL Factory R84 | FC_DL_ClinkerFreeLimeCalc
  功能：融合化学法与在线估算得游离石灰含量，按 ≤1.5% 判合格并给烧成度分级
  开源溯源：无（clean-room 自研，依据公开工艺公式，来源=行业通用公式，许可证=MIT，借鉴点=公式结构）
  规则：R1-R16 全遵守
*)
FUNCTION FC_DL_ClinkerFreeLimeCalc : REAL
VAR_INPUT
    fCaOLabPct : REAL := -1.0; // 化学法实测 f-CaO（负值表示本次无化验值） [%] / lab free lime, negative means not available [%]
    fCaOEstPct : REAL := 1.2; // 在线估算 f-CaO [%] / online estimated free lime [%]
    fLabWeight : REAL := 0.7; // 化验值权重（0~1） [-] / laboratory weight [0,1]
    fLimitPct : REAL := 1.5; // 合格上限 [%] / acceptance limit [%]
    fUnderLoPct : REAL := 0.5; // 过烧判据下限（低于即判过烧） [%] / overburn lower bound [%]
END_VAR
VAR_OUTPUT
    iBurnGrade : INT; // 烧成度分级 0=过烧 1=正常 2=欠烧 [-] / burning grade [-]
    xPass : BOOL; // f-CaO 判合格 [-] / free lime passed [-]
    xValid : BOOL; // 计算结果有效标志 [-] / calculation valid flag [-]
END_VAR
VAR
    fW : REAL; // 实际采用权重（钳位后） [-] / effective weight after clamping [-]
    fCaOPct : REAL; // 融合后 f-CaO [%] / fused free lime [%]
END_VAR

// 段 1｜出口预置（R256）
FC_DL_ClinkerFreeLimeCalc := -1.0; // 哨兵返回 -1（无效） [-] / sentinel return -1, invalid [-]
iBurnGrade := 1; // 分级预置正常 [-] / grade preset to normal [-]
xPass := FALSE; // 合格位预置 FALSE [-] / pass preset false [-]
xValid := FALSE; // 计算完成前不认结果 [-] / unusable before calculation [-]

// 段 2｜非有限拦截 + 域闸（R4/R20）
IF NOT (fCaOLabPct > -1.0E30 AND fCaOLabPct < 1.0E30) OR NOT (fCaOEstPct > -1.0E30 AND fCaOEstPct < 1.0E30) OR NOT (fLabWeight > -1.0E30 AND fLabWeight < 1.0E30) THEN
    RETURN; // 化验值/估算值/权重任一非有限即拒算 [-] / any non finite input rejected [-]
END_IF
IF fCaOEstPct < 0.0 OR NOT (fLimitPct > -1.0E30 AND fLimitPct < 1.0E30) OR NOT (fUnderLoPct > -1.0E30 AND fUnderLoPct < 1.0E30) THEN
    RETURN; // 估算值非负 + 阈值有限闸 [%] / non negative estimate and finite thresholds [%]
END_IF
IF fLimitPct <= 0.0 OR fUnderLoPct < 0.0 OR NOT (fUnderLoPct < fLimitPct) THEN
    RETURN; // 阈值组态闸：0 ≤ 过烧下限 < 合格上限 [%] / threshold config gate [%]
END_IF

// 段 3｜权重钳位与融合（化验值缺失时权重强制归零）
fW := fLabWeight; // 无量纲权重 [-] / dimensionless weight [-]
IF fCaOLabPct < 0.0 THEN
    fW := 0.0; // 无化验值：全部采用在线估算 [-] / no lab value, use the estimate only [-]
END_IF
IF fW > 1.0 THEN
    fW := 1.0; // 权重上限钳位 [-] / clamp the weight high [-]
END_IF
IF fW < 0.0 THEN
    fW := 0.0; // 权重下限钳位 [-] / clamp the weight low [-]
END_IF
IF fW >= 1.0 THEN
    fCaOPct := fCaOLabPct; // 全信化验值 [%] / trust the lab value entirely [%]
ELSE
    fCaOPct := (fCaOLabPct * fW) + (fCaOEstPct * (1.0 - fW)); // % × - + % × - = % / [%] × [-] + [%] × [-] = [%]
END_IF
IF NOT (fCaOPct > -1.0E30 AND fCaOPct < 1.0E30) THEN
    RETURN; // 结果非有限再拦一次 [-] / second finiteness gate [-]
END_IF

// 段 4｜合格判定与烧成度分级（f-CaO 高=欠烧，低=过烧）
IF fCaOPct > fLimitPct THEN
    iBurnGrade := 2; // 欠烧：f-CaO 超上限 [-] / underburnt, free lime above the limit [-]
    xPass := FALSE; // 不合格 [-] / fail [-]
ELSIF fCaOPct < fUnderLoPct THEN
    iBurnGrade := 0; // 过烧：f-CaO 过低（浪费热耗） [-] / overburnt, free lime too low [-]
    xPass := TRUE; // 仍判合格（质量达标，但需节能） [-] / still passing on quality [-]
ELSE
    iBurnGrade := 1; // 正常区间 [-] / normal band [-]
    xPass := TRUE; // 合格 [-] / pass [-]
END_IF
xValid := TRUE; // 链路有效 [-] / chain valid [-]
FC_DL_ClinkerFreeLimeCalc := fCaOPct; // 返回游离石灰 [%] / return the free lime [%]
END_FUNCTION

(* ---- FC_DL_ClinkerLsfCalc.st ---- *)
(*
  DL Factory R84 | FC_DL_ClinkerLsfCalc
  功能：算熟料石灰饱和系数 LSF 并附硅率 SM 与铝率 IM 率值
  开源溯源：无（clean-room 自研，依据公开工艺公式，来源=行业通用公式，许可证=MIT，借鉴点=公式结构）
  规则：R1-R16 全遵守
*)
FUNCTION FC_DL_ClinkerLsfCalc : REAL
VAR_INPUT
    fCaO : REAL := 65.0; // 氧化钙含量 [%] / calcium oxide content [%]
    fSiO2 : REAL := 21.0; // 二氧化硅含量 [%] / silica content [%]
    fAl2O3 : REAL := 5.2; // 三氧化二铝含量 [%] / alumina content [%]
    fFe2O3 : REAL := 3.4; // 三氧化二铁含量 [%] / ferric oxide content [%]
    fLsfLo : REAL := 92.0; // LSF 合格下限 [-] / LSF lower acceptance bound [-]
    fLsfHi : REAL := 98.0; // LSF 合格上限 [-] / LSF upper acceptance bound [-]
END_VAR
VAR_OUTPUT
    fSm : REAL; // 硅率 SM [-] / silica modulus [-]
    fIm : REAL; // 铝率 IM [-] / alumina modulus [-]
    xPass : BOOL; // LSF 落在合格带 [-] / LSF inside the acceptance band [-]
    xValid : BOOL; // 计算结果有效标志 [-] / calculation valid flag [-]
END_VAR
VAR
    fNum : REAL; // LSF 分子（CaO − 1.65Al − 0.35Fe） [%] / LSF numerator [%]
    fLsf : REAL; // LSF 中间量 [-] / LSF intermediate [-]
    fAlFe : REAL; // 铝铁合计（SM 分母） [%] / alumina plus ferric sum [%]
END_VAR

// 段 1｜出口预置（R256）
FC_DL_ClinkerLsfCalc := -1.0; // 哨兵返回 -1（无效） [-] / sentinel return -1, invalid [-]
fSm := 0.0; // 硅率预置零 [-] / silica modulus preset zero [-]
fIm := 0.0; // 铝率预置零 [-] / alumina modulus preset zero [-]
xPass := FALSE; // 合格位预置 FALSE [-] / pass preset false [-]
xValid := FALSE; // 计算完成前不认结果 [-] / unusable before calculation [-]

// 段 2｜非有限拦截 + 域闸（R4/R20）
IF NOT (fCaO > -1.0E30 AND fCaO < 1.0E30) OR NOT (fSiO2 > -1.0E30 AND fSiO2 < 1.0E30) OR NOT (fAl2O3 > -1.0E30 AND fAl2O3 < 1.0E30) OR NOT (fFe2O3 > -1.0E30 AND fFe2O3 < 1.0E30) THEN
    RETURN; // 四项氧化物任一非有限即拒算 [-] / any non finite oxide rejected [-]
END_IF
IF fCaO < 0.0 OR fSiO2 < 1.0E-9 OR fAl2O3 < 0.0 OR fFe2O3 < 1.0E-9 THEN
    RETURN; // SiO2 与 Fe2O3 正域分母闸 + 其余非负闸 [%] / positive denominator gate [%]
END_IF
IF NOT (fLsfLo > -1.0E30 AND fLsfLo < 1.0E30) OR NOT (fLsfHi > -1.0E30 AND fLsfHi < 1.0E30) OR NOT (fLsfLo < fLsfHi) THEN
    RETURN; // 合格带组态闸：下限必须严格小于上限 [-] / acceptance band config gate [-]
END_IF

// 段 3｜LSF = (CaO − 1.65Al2O3 − 0.35Fe2O3) / (2.8 SiO2)
fNum := (fCaO - (1.65 * fAl2O3)) - (0.35 * fFe2O3); // % − % − % = %（系数无量纲） / [%] - [%] - [%] = [%]
fLsf := fNum / (2.8 * fSiO2); // % ÷ % = 无量纲 / [%] / [%] = [-]
IF NOT (fLsf > -1.0E30 AND fLsf < 1.0E30) THEN
    RETURN; // 结果非有限再拦一次 [-] / second finiteness gate [-]
END_IF

// 段 4｜率值：SM = SiO2/(Al+Fe)，IM = Al/Fe
fAlFe := fAl2O3 + fFe2O3; // % + % = % / [%] + [%] = [%]
IF fAlFe < 1.0E-9 THEN
    RETURN; // 分母闸：铝铁合计趋零 [%] / denominator gate on the alumina plus ferric sum [%]
END_IF
fSm := fSiO2 / fAlFe; // % ÷ % = 无量纲 / [%] / [%] = [-]
fIm := fAl2O3 / fFe2O3; // % ÷ % = 无量纲 / [%] / [%] = [-]
IF NOT (fSm > -1.0E30 AND fSm < 1.0E30) OR NOT (fIm > -1.0E30 AND fIm < 1.0E30) THEN
    RETURN; // 率值非有限再拦一次 [-] / second finiteness gate on the moduli [-]
END_IF
xPass := (fLsf >= fLsfLo) AND (fLsf <= fLsfHi); // 带内判据，双边直比 [-] / band verdict with two sided compares [-]
xValid := TRUE; // 链路有效 [-] / chain valid [-]
FC_DL_ClinkerLsfCalc := fLsf; // 返回 LSF [-] / return the LSF [-]
END_FUNCTION

(* ---- FC_DL_CncMrrCalc.st ---- *)
(*
  DL Factory R84 | FC_DL_CncMrrCalc
  功能：算铣削材料去除率 MRR 并折算 cm³/min 与每分钟切屑质量
  开源溯源：无（clean-room 自研，依据公开工艺公式，来源=行业通用公式，许可证=MIT，借鉴点=公式结构）
  规则：R1-R16 全遵守
*)
FUNCTION FC_DL_CncMrrCalc : REAL
VAR_INPUT
    fAp : REAL := 1.0; // 轴向切深 [mm] / axial depth of cut [mm]
    fAe : REAL := 5.0; // 径向切宽 [mm] / radial width of cut [mm]
    fVf : REAL := 800.0; // 进给速度 [mm/min] / feed rate [mm/min]
    fRho : REAL := 7.85; // 材料密度 [g/cm³] / material density [g/cm^3]
END_VAR
VAR_OUTPUT
    fMrrCm3Min : REAL; // 材料去除率折算 [cm³/min] / removal rate in [cm^3/min]
    fChipKgMin : REAL; // 每分钟切屑质量 [kg/min] / chip mass per minute [kg/min]
    xValid : BOOL; // 计算结果有效标志 [-] / calculation valid flag [-]
END_VAR
VAR
    fMrrMm3 : REAL; // 材料去除率原始量 [mm³/min] / raw removal rate [mm^3/min]
    fGramMin : REAL; // 切屑质量流 [g/min] / chip mass flow [g/min]
END_VAR

// 段 1｜出口预置（R256）
FC_DL_CncMrrCalc := -1.0; // 哨兵返回 -1（无效） [-] / sentinel return -1, invalid [-]
fMrrCm3Min := 0.0; // cm³/min 预置零 / preset to zero [cm^3/min]
fChipKgMin := 0.0; // 切屑质量预置零 [kg/min] / chip mass preset zero [kg/min]
xValid := FALSE; // 计算完成前不认结果 [-] / unusable before calculation [-]

// 段 2｜非有限拦截 + 物理域闸（R4/R20）
IF NOT (fAp > -1.0E30 AND fAp < 1.0E30) OR NOT (fAe > -1.0E30 AND fAe < 1.0E30) OR NOT (fVf > -1.0E30 AND fVf < 1.0E30) OR NOT (fRho > -1.0E30 AND fRho < 1.0E30) THEN
    RETURN; // 任一入参为 NaN/Inf 一律拒绝 [-] / any NaN or Inf input rejected [-]
END_IF
IF fAp < 0.0 OR fAe < 0.0 OR fVf < 0.0 THEN
    RETURN; // 几何量与进给不得为负 [-] / geometry and feed must not be negative [-]
END_IF
IF fRho <= 1.0E-9 THEN
    RETURN; // 密度正域闸（避免除零与零质量） [g/cm³] / density positive domain gate [g/cm^3]
END_IF

// 段 3｜主算：MRR = ap × ae × vf
fMrrMm3 := (fAp * fAe) * fVf; // mm × mm × mm/min = mm³/min / [mm] × [mm] × [mm/min] = [mm^3/min]
IF fMrrMm3 <= 0.0 THEN
    RETURN; // 零截面或零进给无去除量 [-] / zero section or zero feed removes nothing [-]
END_IF
fMrrCm3Min := fMrrMm3 / 1000.0; // mm³ ÷ 1000 = cm³（1 cm³ = 1000 mm³） / [mm^3] / 1000 = [cm^3]
fGramMin := fMrrCm3Min * fRho; // cm³/min × g/cm³ = g/min / [cm^3/min] × [g/cm^3] = [g/min]
fChipKgMin := fGramMin / 1000.0; // g/min ÷ 1000 = kg/min / [g/min] / 1000 = [kg/min]
IF NOT (fChipKgMin > -1.0E30 AND fChipKgMin < 1.0E30) THEN
    RETURN; // 结果非有限再拦一次 [-] / second finiteness gate on the result [-]
END_IF
xValid := TRUE; // 链路有效 [-] / chain valid [-]
FC_DL_CncMrrCalc := fMrrMm3; // 返回 MRR [mm³/min] / return the removal rate [mm^3/min]
END_FUNCTION

(* ---- FC_DL_CncSpindleLoadRatio.st ---- *)
(*
  DL Factory R84 | FC_DL_CncSpindleLoadRatio
  功能：算主轴负载率并给过载裕度与 85%/100% 两级报警位
  开源溯源：无（clean-room 自研，依据公开工艺公式，来源=行业通用公式，许可证=MIT，借鉴点=公式结构）
  规则：R1-R16 全遵守
*)
FUNCTION FC_DL_CncSpindleLoadRatio : REAL
VAR_INPUT
    fActualKw : REAL := 0.0; // 主轴实际输出功率 [kW] / actual spindle power [kW]
    fRatedKw : REAL := 7.5; // 主轴额定（连续）功率 [kW] / rated spindle power [kW]
    fWarnPct : REAL := 85.0; // 预警负载率门限 [%] / warning load threshold [%]
    fTripPct : REAL := 100.0; // 停机建议门限 [%] / trip recommendation threshold [%]
END_VAR
VAR_OUTPUT
    fMarginPct : REAL; // 过载裕度（100 − 负载率） [%] / overload margin [%]
    xWarn : BOOL; // 负载率超预警门限 [-] / load above warning threshold [-]
    xTrip : BOOL; // 负载率超停机建议门限 [-] / load above trip threshold [-]
    xValid : BOOL; // 计算结果有效标志 [-] / calculation valid flag [-]
END_VAR
VAR
    fRatioPct : REAL; // 负载率中间量 [%] / load ratio intermediate [%]
END_VAR

// 段 1｜出口预置（R256）
FC_DL_CncSpindleLoadRatio := -1.0; // 哨兵返回 -1（无效） [-] / sentinel return -1, invalid [-]
fMarginPct := 0.0; // 裕度预置零 [%] / margin preset zero [%]
xWarn := FALSE; // 预警位预置 FALSE [-] / warning preset false [-]
xTrip := FALSE; // 停机位预置 FALSE [-] / trip preset false [-]
xValid := FALSE; // 计算完成前不认结果 [-] / unusable before calculation [-]

// 段 2｜非有限拦截 + 额定功率分母闸（R4/R20）
IF NOT (fActualKw > -1.0E30 AND fActualKw < 1.0E30) OR NOT (fRatedKw > -1.0E30 AND fRatedKw < 1.0E30) OR NOT (fWarnPct > -1.0E30 AND fWarnPct < 1.0E30) OR NOT (fTripPct > -1.0E30 AND fTripPct < 1.0E30) THEN
    RETURN; // 任一入参为 NaN/Inf 一律拒绝 [-] / any NaN or Inf input rejected [-]
END_IF
IF fRatedKw < 1.0E-9 THEN
    RETURN; // 额定功率正域分母闸（防除零） [kW] / rated power positive denominator gate [kW]
END_IF
IF NOT (fWarnPct < fTripPct) THEN
    RETURN; // 组态闸：预警门限必须严格小于停机门限 [%] / config gate: warn below trip [%]
END_IF

// 段 3｜主算：负载率 = 实际功率 / 额定功率
fRatioPct := (fActualKw / fRatedKw) * 100.0; // kW ÷ kW × 100 = % / [kW] / [kW] × 100 = [%]
IF NOT (fRatioPct > -1.0E30 AND fRatioPct < 1.0E30) THEN
    RETURN; // 结果非有限再拦一次 [-] / second finiteness gate on the result [-]
END_IF
fMarginPct := 100.0 - fRatioPct; // % − % = %（负值表示已过载） / [%] minus [%] = [%], negative means overloaded
xWarn := fRatioPct > fWarnPct; // 直比门限，禁浮点等值 [-] / direct compare, no float equality [-]
xTrip := fRatioPct > fTripPct; // 直比门限，禁浮点等值 [-] / direct compare, no float equality [-]
xValid := TRUE; // 链路有效 [-] / chain valid [-]
FC_DL_CncSpindleLoadRatio := fRatioPct; // 返回负载率 [%] / return the load ratio [%]
END_FUNCTION

(* ---- FC_DL_CoilWeightEstCalc.st ---- *)
(*
  Name: FC_DL_CoilWeightEstCalc
  Category: DL_Device
  Version: 1.0.0
  Round: R89 / 2026-11-25
  开源溯源：clean-room 自研（族 板带剪切分条卷取，ST 开源生态实测 0 命中，无外部代码引入）
  功能：钢卷重量估算：按带长、带宽、带厚与材料密度算理论重量。
  边界条件：① 四入参全部过非有限闸，任一非有限返回哨兵 -1；
            ② 负值与零值一律剔除（长度 ≤ 0、宽厚 ≤ 0 视为无料），返回哨兵 -1，不静默输出 0 kg；
            ③ 尺寸与密度按工程域闸限定，密度取钢 7000~8000 kg/m3 带宽区间含不锈钢与碳钢。
  量纲自证：L[m] × W[m] × T[m] = m3；m3 × ρ[kg/m3] = kg。
*)
FUNCTION FC_DL_CoilWeightEstCalc : REAL
VAR_INPUT
    fLengthM : REAL;        (* 带长 [m] Strip length [m] *)
    fWidthMm : REAL;        (* 带宽 [mm] Strip width [mm] *)
    fThkMm : REAL;          (* 带厚 [mm] Strip thickness [mm] *)
    fDensityKgM3 : REAL;    (* 材料密度 [kg/m3] Material density [kg/m3] *)
END_VAR
VAR_OUTPUT
    fWeightKg : REAL;       (* 钢卷重量 [kg] Coil weight [kg] *)
    xValid : BOOL;          (* 计算有效性标志 [-] Calculation valid flag *)
END_VAR
VAR CONSTANT
    DL_EPS : REAL := 1.0E-9;        (* 判据容差 [-] Criterion tolerance *)
    DL_MM_TO_M : REAL := 1000.0;    (* 毫米 → 米换算 [mm/m] Millimetre to metre *)
    DL_L_MAX : REAL := 100000.0;    (* 带长上限 [m] Length ceiling [m] *)
    DL_W_MIN : REAL := 100.0;       (* 带宽下限 [mm] Width floor [mm] *)
    DL_W_MAX : REAL := 2500.0;      (* 带宽上限 [mm] Width ceiling [mm] *)
    DL_T_MIN : REAL := 0.05;        (* 带厚下限 [mm] Thickness floor [mm] *)
    DL_T_MAX : REAL := 12.0;        (* 带厚上限 [mm] Thickness ceiling [mm] *)
    DL_RHO_MIN : REAL := 7000.0;    (* 密度下限 [kg/m3] Density floor [kg/m3] *)
    DL_RHO_MAX : REAL := 8000.0;    (* 密度上限 [kg/m3] Density ceiling [kg/m3] *)
END_VAR
VAR
    fVolM3 : REAL;  (* 带钢体积 [m3] Strip volume [m3] *)
END_VAR
(* 出口预置：两出口统一预置（R256） *)
fWeightKg := 0.0; xValid := FALSE;
(* 非有限闸：NaN 自反判 + Inf 差值自减判，四入参全枚举 *)
IF (fLengthM <> fLengthM) OR ((fLengthM - fLengthM) <> 0.0)
   OR (fWidthMm <> fWidthMm) OR ((fWidthMm - fWidthMm) <> 0.0)
   OR (fThkMm <> fThkMm) OR ((fThkMm - fThkMm) <> 0.0)
   OR (fDensityKgM3 <> fDensityKgM3) OR ((fDensityKgM3 - fDensityKgM3) <> 0.0) THEN
    FC_DL_CoilWeightEstCalc := -1.0;        (* 哨兵 -1：入参非有限 / Sentinel -1, non-finite input *)
    RETURN;
END_IF
(* 组态域闸：零与负值一律剔除，尺寸与密度按工程域限定 *)
IF (fLengthM <= DL_EPS) OR (fLengthM > DL_L_MAX)
   OR (fWidthMm < DL_W_MIN) OR (fWidthMm > DL_W_MAX)
   OR (fThkMm < DL_T_MIN) OR (fThkMm > DL_T_MAX)
   OR (fDensityKgM3 < DL_RHO_MIN) OR (fDensityKgM3 > DL_RHO_MAX) THEN
    FC_DL_CoilWeightEstCalc := -1.0;        (* 哨兵 -1：无料或越域 / Sentinel -1, no material or out of range *)
    RETURN;
END_IF
(* 体积：mm → m 后三向相乘，量纲 m3 *)
fVolM3 := fLengthM * (fWidthMm / DL_MM_TO_M) * (fThkMm / DL_MM_TO_M);
(* 重量：m3 × kg/m3 = kg *)
fWeightKg := fVolM3 * fDensityKgM3;
xValid := TRUE;                             (* 链路有效 / Chain valid *)
FC_DL_CoilWeightEstCalc := fWeightKg;
END_FUNCTION

(* ---- FC_DL_ComponentRulEstimate.st ---- *)
(*
  道莅工业代码库 / Daoli Industrial ST Library
  组件: FC_DL_ComponentRulEstimate
  分类: DL_Device
  开源溯源: 无（clean-room 工程公式自研；参考公开工艺计算公式，未复制任何受版权保护代码）
  许可证: 本项目自有 (MIT)
  功能: 依据健康度两次采样外推退化斜率与剩余寿命 RUL，并判定退化加速
*)
FUNCTION FC_DL_ComponentRulEstimate : BOOL
VAR_INPUT
    rHealthNow : REAL; // 本次健康度采样 [%]，100 = 全新 / current health sample in percent, 100 is new
    rHealthPrev : REAL; // 上次健康度采样 [%] / previous health sample
    rHoursDelta : REAL; // 两次采样间隔运行小时 [h] / operating hours between samples
    rFailThr : REAL; // 失效门限健康度 [%] / failure threshold health
END_VAR
VAR_OUTPUT
    rRulHours : REAL; // 剩余寿命 [h]，上限哨兵 99999 / remaining useful life, sentinel 99999
    rSlopePerH : REAL; // 退化斜率 [%/h] / degradation slope
    bValid : BOOL; // 结果有效位 [-] / result valid flag
    bAccel : BOOL; // 退化加速标志（斜率低于 -0.001 %/h）[-] / accelerated degradation flag
    iErrCode : INT; // 事件码 0=正常 1=间隔非法 2=无退化（哨兵寿命）3=已到门限 4=结果非有限 / event code
END_VAR
VAR CONSTANT
    rSlopeDead : REAL := 1.0E-9; // 斜率死区（视作无退化）[%/h] / slope dead band
    rSlopeAccel : REAL := -0.001; // 加速退化判据斜率 [%/h] / accelerated degradation slope threshold
    rRulCap : REAL := 99999.0; // 剩余寿命上限哨兵 [h] / remaining life sentinel cap
END_VAR
VAR
    rSlopeRaw : REAL; // 未限幅斜率 [%/h] / unchecked slope
    rRulRaw : REAL; // 未限幅剩余寿命 [h] / unchecked remaining life
    rHeadRoom : REAL; // 剩余健康度余量 [%] / health headroom
END_VAR

    // —— 段 0：全路径预清 —— //
    rSlopeRaw := 0.0;
    rRulRaw := 0.0;
    rHeadRoom := 0.0;
    rRulHours := 0.0;
    rSlopePerH := 0.0;
    bValid := FALSE;
    bAccel := FALSE;
    iErrCode := 0;
    FC_DL_ComponentRulEstimate := FALSE;
    // —— 段 1：分母闸（采样间隔必须为正） —— //
    IF rHoursDelta <= 0.0 THEN
        iErrCode := 1; // 采样间隔非法，斜率无定义 / invalid interval, slope undefined
        RETURN;
    END_IF;
    // —— 段 2：量纲链 (% - %)/(h) = %/h —— //
    rSlopeRaw := (rHealthNow - rHealthPrev) / rHoursDelta; // 退化斜率 [%/h] / degradation slope
    IF ABS(rSlopeRaw) > 1.0E15 THEN
        iErrCode := 4; // 结果非有限，强制归零 / non-finite result, forced to zero
        RETURN;
    END_IF;
    rSlopePerH := rSlopeRaw;
    // —— 段 3：无退化判据（死区内视作零斜率，寿命取哨兵） —— //
    IF ABS(rSlopePerH) < rSlopeDead THEN
        rRulHours := rRulCap; // 哨兵寿命 [h] / sentinel life
        iErrCode := 2; // 信息级：无退化 / info level: no degradation
        bValid := TRUE;
        FC_DL_ComponentRulEstimate := TRUE;
        RETURN;
    END_IF;
    // —— 段 4：剩余健康度余量与 RUL（分母闸：|斜率| 已过死区） —— //
    rHeadRoom := rHealthNow - rFailThr; // 剩余健康度 [%] / health headroom
    IF rHeadRoom <= 0.0 THEN
        rRulHours := 0.0; // 已到或越过失效门限 / threshold already reached
        iErrCode := 3; // 信息级：寿命耗尽 / info level: life exhausted
        bAccel := rSlopePerH < rSlopeAccel; // 仍给出加速判据 / acceleration still reported
        bValid := TRUE;
        FC_DL_ComponentRulEstimate := TRUE;
        RETURN;
    END_IF;
    rRulRaw := rHeadRoom / ABS(rSlopePerH); // 量纲 %/(%/h) = h / remaining life in hours
    IF ABS(rRulRaw) > 1.0E15 THEN
        rRulHours := 0.0;
        iErrCode := 4; // 结果非有限，强制归零 / non-finite result, forced to zero
        RETURN;
    END_IF;
    IF rRulRaw > rRulCap THEN
        rRulHours := rRulCap; // 上限饱和 / saturate at cap
    ELSE
        rRulHours := rRulRaw;
    END_IF;
    bAccel := rSlopePerH < rSlopeAccel; // 退化加速标志 [-] / accelerated degradation flag
    bValid := TRUE;
    FC_DL_ComponentRulEstimate := TRUE;
END_FUNCTION

(* ---- FC_DL_CoolantConcCalc.st ---- *)
(*
  DL Factory R84 | FC_DL_CoolantConcCalc
  功能：由折光读数算切削液浓度，并按两液混合守恒算补原液量与补水量
  开源溯源：无（clean-room 自研，依据公开工艺公式，来源=行业通用公式，许可证=MIT，借鉴点=公式结构）
  规则：R1-R16 全遵守
*)
FUNCTION FC_DL_CoolantConcCalc : REAL
VAR_INPUT
    fRefractBrix : REAL := 3.0; // 折光仪读数（Brix 刻度） [%] / refractometer reading [%]
    fRefractCoef : REAL := 2.0; // 折光换算系数（无量纲） [-] / refractometer conversion factor [-]
    fVolL : REAL := 500.0; // 当前槽液体积 [L] / current sump volume [L]
    fTargetPct : REAL := 8.0; // 目标工作浓度 [%] / target working concentration [%]
END_VAR
VAR_OUTPUT
    fAddConcL : REAL; // 需补原液体积 [L] / raw concentrate to add [L]
    fAddWaterL : REAL; // 需补清水体积 [L] / water to add [L]
    xValid : BOOL; // 计算结果有效标志 [-] / calculation valid flag [-]
END_VAR
VAR
    fCurPct : REAL; // 当前实测浓度 [%] / measured concentration [%]
    fDen : REAL; // 混合守恒分母（无量纲/百分比项） [-] / conservation denominator [-]
END_VAR

// 段 1｜出口预置（R256）
FC_DL_CoolantConcCalc := -1.0; // 哨兵返回 -1（无效） [-] / sentinel return -1, invalid [-]
fAddConcL := 0.0; // 补原液预置零 [L] / concentrate preset zero [L]
fAddWaterL := 0.0; // 补水预置零 [L] / water preset zero [L]
xValid := FALSE; // 计算完成前不认结果 [-] / unusable before calculation [-]

// 段 2｜非有限拦截 + 域闸（R4/R20）
IF NOT (fRefractBrix > -1.0E30 AND fRefractBrix < 1.0E30) OR NOT (fRefractCoef > -1.0E30 AND fRefractCoef < 1.0E30) OR NOT (fVolL > -1.0E30 AND fVolL < 1.0E30) OR NOT (fTargetPct > -1.0E30 AND fTargetPct < 1.0E30) THEN
    RETURN; // 任一入参为 NaN/Inf 一律拒绝 [-] / any NaN or Inf input rejected [-]
END_IF
IF fRefractCoef < 1.0E-9 OR fVolL < 0.0 OR fTargetPct < 1.0E-9 OR fTargetPct > 99.0 THEN
    RETURN; // 系数/体积/目标浓度域闸（含除零防护） [%/L] / factor, volume and target domain gate [%/L]
END_IF

// 段 3｜当前浓度 = 折光读数 × 折光系数
fCurPct := fRefractBrix * fRefractCoef; // % × 无量纲 = % / [%] × [-] = [%]

// 段 4｜两液混合守恒：原液按 100% 计，水按 0% 计
IF fCurPct < fTargetPct THEN
    fDen := 100.0 - fTargetPct; // 100% − 目标% = 百分点 / [%] minus [%] = [%]
    IF fDen < 1.0E-9 THEN
        RETURN; // 分母闸：目标浓度逼近 100% 无解 [%] / denominator gate near 100 [%]
    END_IF
    fAddConcL := (fVolL * (fTargetPct - fCurPct)) / fDen; // L × % ÷ % = L（守恒：V·c + 100·a = t·(V+a)） / [L] × [%] / [%] = [L]
    fAddWaterL := 0.0; // 浓度偏低不补水 [L] / no water while low [L]
ELSE
    IF fTargetPct < 1.0E-9 THEN
        RETURN; // 分母闸：目标浓度趋零 [%] / denominator gate on zero target [%]
    END_IF
    fAddWaterL := (fVolL * (fCurPct - fTargetPct)) / fTargetPct; // L × % ÷ % = L（守恒：V·c = t·(V+w)） / [L] × [%] / [%] = [L]
    fAddConcL := 0.0; // 浓度偏高不补原液 [L] / no concentrate while high [L]
END_IF
IF NOT (fAddConcL > -1.0E30 AND fAddConcL < 1.0E30) OR NOT (fAddWaterL > -1.0E30 AND fAddWaterL < 1.0E30) THEN
    RETURN; // 结果非有限再拦一次 [-] / second finiteness gate on the results [-]
END_IF
xValid := TRUE; // 链路有效 [-] / chain valid [-]
FC_DL_CoolantConcCalc := fCurPct; // 返回当前浓度 [%] / return the measured concentration [%]
END_FUNCTION

(* ---- FC_DL_CrahCoolingCapacityCalc.st ---- *)
(*
 * FC_DL_CrahCoolingCapacityCalc | C2 | DL_Device
 * 功能：精密空调显热制冷量（按风量、送回风温差与空气物性）       单位：风量 [m³/h]、温差 [K]、密度 [kg/m³]、比热 [kJ/(kg·K)]、制冷量 [kW]
 * 工况边界：适用于干工况显热计算（不含潜热与风机温升）；风量、密度、比热须 >0 且有限，回风温度须高于送风温度，否则制冷量按 0 发布并置 xValid=FALSE；ρ、cp 取标准空气 1.2 / 1.005，高原或高温工况须现场修正
 * 代数值回代：V=8000 m³/h、ΔT=13 K、ρ=1.2、cp=1.005 → 1.2×1.005×2.2222×13=34.83 kW（spec 记 34.8 kW，一致）
 * 开源溯源：clean-room 自研，未复制任何第三方代码（无外部来源）
 *)
FUNCTION FC_DL_CrahCoolingCapacityCalc : BOOL
VAR_INPUT
    rAirflowM3h : REAL := 8000.0;    // 送风量 | supply air volume flow [m³/h]
    rTreturnC   : REAL := 35.0;      // 回风温度 | return air temperature [℃]
    rTsupplyC   : REAL := 22.0;      // 送风温度 | supply air temperature [℃]
    rRho        : REAL := 1.2;       // 空气密度 | air density [kg/m³]
    rCp         : REAL := 1.005;     // 空气定压比热 | air specific heat at constant pressure [kJ/(kg·K)]
END_VAR
VAR_OUTPUT
    rCoolingKw : REAL;               // 显热制冷量 | sensible cooling capacity [kW]
    rDeltaTK   : REAL;               // 送回风温差 | return to supply temperature difference [K]
    rMassFlowKgs : REAL;             // 空气质量流量 | air mass flow [kg/s]
    xValid     : BOOL;               // 输出有效 | outputs valid
END_VAR
VAR
    xFinV   : BOOL;                  // 风量有限性 | airflow is finite
    xFinTr  : BOOL;                  // 回风温度有限性 | return temperature is finite
    xFinTs  : BOOL;                  // 送风温度有限性 | supply temperature is finite
    xFinRho : BOOL;                  // 密度有限性 | density is finite
    xFinCp  : BOOL;                  // 比热有限性 | specific heat is finite
    rVolM3s : REAL;                  // 体积流量（m³/s）| volume flow in SI units [m³/s]
END_VAR
VAR CONSTANT
    DL_CCC_SEC_PER_HOUR : REAL := 3600.0;   // 小时转秒系数 | hours to seconds factor [s/h]
END_VAR

// 段1｜非有限闸（R19）
xFinV := (rAirflowM3h = rAirflowM3h) AND ((rAirflowM3h - rAirflowM3h) = 0.0);
xFinTr := (rTreturnC = rTreturnC) AND ((rTreturnC - rTreturnC) = 0.0);
xFinTs := (rTsupplyC = rTsupplyC) AND ((rTsupplyC - rTsupplyC) = 0.0);
xFinRho := (rRho = rRho) AND ((rRho - rRho) = 0.0);
xFinCp := (rCp = rCp) AND ((rCp - rCp) = 0.0);
IF (NOT xFinV) OR (NOT xFinTr) OR (NOT xFinTs) OR (NOT xFinRho) OR (NOT xFinCp) THEN
    rCoolingKw := 0.0;               // 安全值：制冷量 0 | safe value, zero capacity
    rDeltaTK := 0.0;
    rMassFlowKgs := 0.0;
    xValid := FALSE;
    FC_DL_CrahCoolingCapacityCalc := FALSE;
    RETURN;
END_IF

// 段2｜域闸：风量/密度/比热须为正（均入乘积链），回风须高于送风
IF (rAirflowM3h <= 0.0) OR (rRho <= 0.0) OR (rCp <= 0.0) OR (rTreturnC <= rTsupplyC) THEN
    rCoolingKw := 0.0;
    rDeltaTK := 0.0;
    rMassFlowKgs := 0.0;
    xValid := FALSE;
    FC_DL_CrahCoolingCapacityCalc := FALSE;
    RETURN;
END_IF

// 段3｜算法：Q_kW = ρ×cp×V(m³/s)×ΔT
rDeltaTK := rTreturnC - rTsupplyC;
rVolM3s := rAirflowM3h / DL_CCC_SEC_PER_HOUR;
rMassFlowKgs := rRho * rVolM3s;
rCoolingKw := rMassFlowKgs * rCp * rDeltaTK;

// 段4｜出口
xValid := TRUE;
FC_DL_CrahCoolingCapacityCalc := TRUE;
END_FUNCTION

(* ---- FC_DL_CrahSupplyTempResetCalc.st ---- *)
(*
 * FC_DL_CrahSupplyTempResetCalc | C2 | DL_Device
 * 功能：按最不利机柜进风温度重置精密空调送风温度设定值       单位：温度 [℃]、增益 [1]
 * 工况边界：单回路比例重置，适用于机柜进风温度反馈可信（无传感器故障）场合；上下限须满足 min<max 且增益 ≥0，否则 xValid=FALSE 并输出下限安全值；clamped 判定以未钳位的原始计算值为准（R24，禁止先夹再判）
 * 代数值回代：worst=27、target=24、gain=0.6、base=20、限 [18,27] → sp=20+0.6×3=21.8 ℃，未打限幅 → xClamped=FALSE（与 spec 回代行一致）
 * 开源溯源：clean-room 自研，未复制任何第三方代码（无外部来源）
 *)
FUNCTION FC_DL_CrahSupplyTempResetCalc : BOOL
VAR_INPUT
    rWorstRackInletC : REAL := 27.0;  // 最不利机柜进风温度 | worst rack inlet temperature [℃]
    rRackTargetC     : REAL := 24.0;  // 机柜进风目标温度 | rack inlet target temperature [℃]
    rGain            : REAL := 0.6;   // 重置增益 | reset gain [1]
    rMinC            : REAL := 18.0;  // 送风设定下限 | supply setpoint lower limit [℃]
    rMaxC            : REAL := 27.0;  // 送风设定上限 | supply setpoint upper limit [℃]
    rBaseC           : REAL := 20.0;  // 基准送风温度 | base supply temperature [℃]
END_VAR
VAR_OUTPUT
    rSupplySetpointC : REAL;          // 送风温度设定值 | supply temperature setpoint [℃]
    rRawSetpointC    : REAL;          // 未钳位的原始计算值 | raw setpoint before clamping [℃]
    xClamped         : BOOL;          // 已打限幅（信息级）| clamped against the limits, informational
    xValid           : BOOL;          // 输出有效 | outputs valid
END_VAR
VAR
    xFinWorst : BOOL;                 // 最不利温度有限性 | worst temperature is finite
    xFinTg    : BOOL;                 // 目标温度有限性 | target temperature is finite
    xFinGain  : BOOL;                 // 增益有限性 | gain is finite
    xFinMin   : BOOL;                 // 下限有限性 | lower limit is finite
    xFinMax   : BOOL;                 // 上限有限性 | upper limit is finite
    xFinBase  : BOOL;                 // 基准有限性 | base temperature is finite
END_VAR
VAR CONSTANT
    DL_CSR_EPS : REAL := 1.0E-6;      // 浮点比较容差 | floating comparison tolerance [℃]
END_VAR

// 段1｜非有限闸（R19：非有限即输出下限安全值，避免 NaN 流入设定值）
xFinWorst := (rWorstRackInletC = rWorstRackInletC) AND ((rWorstRackInletC - rWorstRackInletC) = 0.0);
xFinTg := (rRackTargetC = rRackTargetC) AND ((rRackTargetC - rRackTargetC) = 0.0);
xFinGain := (rGain = rGain) AND ((rGain - rGain) = 0.0);
xFinMin := (rMinC = rMinC) AND ((rMinC - rMinC) = 0.0);
xFinMax := (rMaxC = rMaxC) AND ((rMaxC - rMaxC) = 0.0);
xFinBase := (rBaseC = rBaseC) AND ((rBaseC - rBaseC) = 0.0);
IF (NOT xFinWorst) OR (NOT xFinTg) OR (NOT xFinGain) OR (NOT xFinMin)
   OR (NOT xFinMax) OR (NOT xFinBase) THEN
    rSupplySetpointC := 18.0;        // 安全值：取下限（不结露的保守侧）| safe value, the conservative lower limit
    rRawSetpointC := 18.0;
    xClamped := TRUE;
    xValid := FALSE;
    FC_DL_CrahSupplyTempResetCalc := FALSE;
    RETURN;
END_IF

// 段2｜域闸：限幅区间有效且增益非负
IF (rMaxC <= rMinC) OR (rGain < 0.0) THEN
    rSupplySetpointC := rMinC;       // 安全值：取下限 | safe value, the lower limit
    rRawSetpointC := rMinC;
    xClamped := TRUE;
    xValid := FALSE;
    FC_DL_CrahSupplyTempResetCalc := FALSE;
    RETURN;
END_IF

// 段3｜算法：sp = base + gain×(worst − target)
rRawSetpointC := rBaseC + rGain * (rWorstRackInletC - rRackTargetC);

// 段4｜限幅与打限标志（判据取自未钳位原始值，R24）
xClamped := (rRawSetpointC > (rMaxC + DL_CSR_EPS)) OR (rRawSetpointC < (rMinC - DL_CSR_EPS));
rSupplySetpointC := LIMIT(rMinC, rRawSetpointC, rMaxC);

// 段5｜出口
xValid := TRUE;
FC_DL_CrahSupplyTempResetCalc := TRUE;
END_FUNCTION

(* ---- FC_DL_CraneWindSpeedLimitChk.st ---- *)
(*
 * FC_DL_CraneWindSpeedLimitChk | C1 | DL_Device
 * 功能：风速分级作业限幅判定（正常 / 降速 / 停工 / 锚定）       单位：风速 [m/s]，分级与许可为枚举码与布尔
 * 工况边界：阈值取 GB/T 3811 工作状态风 13.8 / 20.0 / 25.0 m/s；判据以 MAX(3 s 均值, 阵风) 为最不利值；风速 NaN/Inf 或超 40 m/s 量程一律按锚定侧安全值输出；本件不含滞环，滞环由序列 FB 承担
 * 代数值回代：MAX(均值,阵风)=22.0 → nLevel=2（20~25 停工）；26.0 → nLevel=3（锚定）；8.0 → nLevel=0（正常）（与 spec 回代行一致）
 * 开源溯源：clean-room 自研，未复制任何第三方代码（无外部来源）
 *)
FUNCTION FC_DL_CraneWindSpeedLimitChk : BOOL
VAR_INPUT
    rWindMs : REAL;                  // 风速 3 s 均值 | wind speed, 3 s mean [m/s]
    rGustMs : REAL;                  // 风速阵风值（3 s 均值窗内的最大瞬时）| gust value within the 3 s window [m/s]
END_VAR
VAR_OUTPUT
    nLevel         : INT;            // 0=正常 / 1=降速 / 2=停工 / 3=锚定 | 0 normal, 1 derate, 2 stop, 3 anchor
    xPermitWork    : BOOL;           // 允许作业 | work permitted
    xPermitTravel  : BOOL;           // 允许行车 | travelling permitted
    xRequireAnchor : BOOL;           // 要求锚定 | anchoring required
    xPermitFullSpeed : BOOL;         // 允许全速（仅 0 级）| full speed permitted, level 0 only
    xValid         : BOOL;           // 输出有效（风速可信）| outputs valid, the wind reading is trustworthy
END_VAR
VAR
    xFinMean : BOOL;                 // 均值有限性 | mean value is finite
    xFinGust : BOOL;                 // 阵风有限性 | gust value is finite
    rWindChk : REAL;                 // 判定用风速（取均值与阵风的较大者）| wind used for grading, the worse of the two
END_VAR
VAR CONSTANT
    DL_CWS_DERATE : REAL := 13.8;    // 降速阈 | derating threshold [m/s]
    DL_CWS_STOP   : REAL := 20.0;    // 停工阈 | stop threshold [m/s]
    DL_CWS_ANCHOR : REAL := 25.0;    // 锚定阈 | anchoring threshold [m/s]
    DL_CWS_MAX    : REAL := 40.0;    // 风速量程上限 | upper wind range limit [m/s]
END_VAR

// 段1｜非有限闸（R19：不可信即按锚定侧安全值输出，不让非有限值参与比较）
xFinMean := (rWindMs = rWindMs) AND ((rWindMs - rWindMs) = 0.0);
xFinGust := (rGustMs = rGustMs) AND ((rGustMs - rGustMs) = 0.0);
IF (NOT xFinMean) OR (NOT xFinGust) THEN
    nLevel := 3;                     // 安全值：最高级（锚定）| safe value, the highest level
    xPermitWork := FALSE;
    xPermitTravel := FALSE;
    xRequireAnchor := TRUE;
    xPermitFullSpeed := FALSE;
    xValid := FALSE;
    FC_DL_CraneWindSpeedLimitChk := FALSE;
    RETURN;
END_IF

// 段2｜域闸：负风速或超量程同样按不可信处理（判据与出口同源，R24）
IF (rWindMs < 0.0) OR (rGustMs < 0.0) OR (rWindMs > DL_CWS_MAX) OR (rGustMs > DL_CWS_MAX) THEN
    nLevel := 3;
    xPermitWork := FALSE;
    xPermitTravel := FALSE;
    xRequireAnchor := TRUE;
    xPermitFullSpeed := FALSE;
    xValid := FALSE;
    FC_DL_CraneWindSpeedLimitChk := FALSE;
    RETURN;
END_IF

// 段3｜算法：以最不利值（均值与阵风的较大者）分级
rWindChk := MAX(rWindMs, rGustMs);
nLevel := 0;
xPermitWork := TRUE;
xPermitTravel := TRUE;
xRequireAnchor := FALSE;
xPermitFullSpeed := TRUE;
IF rWindChk > DL_CWS_ANCHOR THEN
    nLevel := 3;                     // >25：锚定 | above 25, anchor
    xPermitWork := FALSE;
    xPermitTravel := FALSE;
    xRequireAnchor := TRUE;
    xPermitFullSpeed := FALSE;
ELSIF rWindChk > DL_CWS_STOP THEN
    nLevel := 2;                     // 20~25：停工 | 20 to 25, stop
    xPermitWork := FALSE;
    xPermitTravel := FALSE;
    xRequireAnchor := FALSE;
    xPermitFullSpeed := FALSE;
ELSIF rWindChk >= DL_CWS_DERATE THEN
    nLevel := 1;                     // 13.8~20：降速作业 | 13.8 to 20, derated working
    xPermitWork := TRUE;
    xPermitTravel := TRUE;
    xRequireAnchor := FALSE;
    xPermitFullSpeed := FALSE;
END_IF

// 段4｜出口
xValid := TRUE;
FC_DL_CraneWindSpeedLimitChk := TRUE;
END_FUNCTION

(* ---- FC_DL_CuttingForceCalc.st ---- *)
(*
  DL Factory R84 | FC_DL_CuttingForceCalc
  功能：按比切削力模型算车削主切削力 Fc 与单位切削功率 Pc
  开源溯源：无（clean-room 自研，依据公开工艺公式，来源=行业通用公式，许可证=MIT，借鉴点=公式结构）
  规则：R1-R16 全遵守
*)
FUNCTION FC_DL_CuttingForceCalc : REAL
VAR_INPUT
    fKc : REAL := 2000.0; // 材料比切削力 [N/mm²] / specific cutting force [N/mm^2]
    fAp : REAL := 1.0; // 背吃刀量（切深） [mm] / depth of cut [mm]
    fFeed : REAL := 0.2; // 每转进给量 [mm/r] / feed per revolution [mm/rev]
    fVc : REAL := 150.0; // 切削线速度 [m/min] / cutting speed [m/min]
    fKcRef : REAL := 1.0; // 比切削力修正系数（无量纲） [-] / specific force correction factor [-]
END_VAR
VAR_OUTPUT
    fUnitPowerKw : REAL; // 单位切削功率 [kW] / unit cutting power [kW]
    xValid : BOOL; // 计算结果有效标志 [-] / calculation valid flag [-]
END_VAR
VAR
    fKcEff : REAL; // 修正后比切削力 [N/mm²] / corrected specific cutting force [N/mm^2]
    fFcRaw : REAL; // 切削力中间量 [N] / cutting force intermediate [N]
END_VAR

// 段 1｜出口预置（R256）
FC_DL_CuttingForceCalc := -1.0; // 哨兵返回 -1（无效） [-] / sentinel return -1, invalid [-]
fUnitPowerKw := 0.0; // 功率预置零 [kW] / power preset to zero [kW]
xValid := FALSE; // 计算完成前不认结果 [-] / unusable before calculation [-]

// 段 2｜非有限拦截 + 物理域闸（R4/R20）
IF NOT (fKc > -1.0E30 AND fKc < 1.0E30) OR NOT (fAp > -1.0E30 AND fAp < 1.0E30) OR NOT (fFeed > -1.0E30 AND fFeed < 1.0E30) OR NOT (fVc > -1.0E30 AND fVc < 1.0E30) OR NOT (fKcRef > -1.0E30 AND fKcRef < 1.0E30) THEN
    RETURN; // 任一入参为 NaN/Inf 一律拒绝 [-] / any NaN or Inf input rejected [-]
END_IF
IF fKc <= 0.0 OR fAp < 0.0 OR fFeed < 0.0 OR fVc < 0.0 THEN
    RETURN; // 比切削力非正或几何量为负即非法 [-] / non positive force or negative geometry [-]
END_IF
IF ABS(fKcRef) < 1.0E-9 THEN
    RETURN; // 分母闸：修正系数趋零 [-] / denominator gate on correction factor [-]
END_IF

// 段 3｜主算：Fc 与 Pc
fKcEff := fKc / fKcRef; // N/mm² ÷ 无量纲 = N/mm² / [N/mm^2] divided by [-]
fFcRaw := (fKcEff * fAp) * fFeed; // N/mm² × mm × mm/r = N（切屑截面积按每转计） / [N/mm^2] × mm × mm/rev = N
IF fFcRaw <= 0.0 THEN
    RETURN; // 零切深或零进给无切削意义 [-] / zero depth or zero feed carries no cut [-]
END_IF
fUnitPowerKw := fFcRaw * fVc / 60000.0; // N × m/min ÷ 60000 = kW（60000 = 60 s × 1000 W） / [N] × [m/min] / 60000 = kW
IF NOT (fUnitPowerKw > -1.0E30 AND fUnitPowerKw < 1.0E30) THEN
    RETURN; // 结果非有限再拦一次 [-] / second finiteness gate on the result [-]
END_IF
xValid := TRUE; // 链路有效 [-] / chain valid [-]
FC_DL_CuttingForceCalc := fFcRaw; // 返回主切削力 [N] / return the cutting force [N]
END_FUNCTION

(* ---- FC_DL_DelubeResidualCarbonCalc.st ---- *)
(*
  Component : FC_DL_DelubeResidualCarbonCalc
  Category  : DL_Device
  Type      : FC
  Complexity: C2
  VERSION   : v1.0.0
  功能      : 润滑剂烧除残碳估算：按烧除区露点、温度与停留时间三个修正因子折算残碳百分比，并与限值比较给出合格判定。
  开源溯源  : 道莅原创 clean-room 自研（无外部代码引用）｜License: MIT
  边界条件  : ① 三个基准量（露点、温度、停留时间）须 > 1e-9，否则返回哨兵 -1；
              ② 各修正因子双侧钳位 0.5~2.0，防单因子离群拉爆残碳估算；
              ③ 露点越高、温度越低、停留越短则残碳越高（三者方向各不相同，逐项显式建模）。
*)
FUNCTION FC_DL_DelubeResidualCarbonCalc : REAL
VAR_INPUT
    fLubePct     : REAL;   (* 润滑剂添加量 [%] Lubricant content *)
    fDewPointC   : REAL;   (* 烧除区露点 [°C] Delube zone dew point *)
    fZoneTempC   : REAL;   (* 烧除区温度 [°C] Delube zone temperature *)
    fResidTimeMin: REAL;   (* 烧除区停留时间 [min] Delube zone residence time *)
    fDewRefC     : REAL;   (* 露点基准 [°C] Dew point reference *)
    fTempRefC    : REAL;   (* 温度基准 [°C] Temperature reference *)
    fTimeRefMin  : REAL;   (* 停留时间基准 [min] Residence time reference *)
    fLimitPct    : REAL;   (* 残碳合格限 [%] Residual carbon limit *)
END_VAR
VAR_OUTPUT
    fResidualPct : REAL;  (* 残碳估算值 [%] Estimated residual carbon *)
    fKCoef       : REAL;  (* 综合修正系数 [-] Composite correction coefficient *)
    xQualified   : BOOL;  (* 残碳合格标志 [-] Residual carbon qualified flag *)
    xValid       : BOOL;  (* 计算有效性标志 [-] Calculation valid flag *)
END_VAR
VAR CONSTANT
    DL_EPS      : REAL := 1.0E-9;   (* 除零判定容差 [无量纲] Divide-by-zero tolerance *)
    DL_K_MIN    : REAL := 0.5;      (* 修正因子下限 [-] Correction factor lower clamp *)
    DL_K_MAX    : REAL := 2.0;      (* 修正因子上限 [-] Correction factor upper clamp *)
    DL_DEW_K    : REAL := 0.02;     (* 露点修正斜率 [1/°C] Dew point slope *)
    DL_TMP_K    : REAL := 0.002;    (* 温度修正斜率 [1/°C] Temperature slope *)
    DL_ZERO     : REAL := 0.0;      (* 零常量 [无量纲] Zero constant *)
END_VAR
VAR
    fKDew  : REAL;   (* 露点修正因子 [-] Dew point factor *)
    fKTmp  : REAL;   (* 温度修正因子 [-] Temperature factor *)
    fKTime : REAL;   (* 停留时间修正因子 [-] Residence time factor *)
END_VAR
(* 出口预置：四出口统一预置 *)
fResidualPct := 0.0; fKCoef := 1.0; xQualified := FALSE; xValid := FALSE;
(* 非有限拦截：自反判 NaN，自身差值判 Inf *)
IF (fLubePct <> fLubePct) OR ((fLubePct - fLubePct) <> 0.0)
   OR (fDewPointC <> fDewPointC) OR ((fDewPointC - fDewPointC) <> 0.0)
   OR (fZoneTempC <> fZoneTempC) OR ((fZoneTempC - fZoneTempC) <> 0.0)
   OR (fResidTimeMin <> fResidTimeMin) OR ((fResidTimeMin - fResidTimeMin) <> 0.0)
   OR (fDewRefC <> fDewRefC) OR ((fDewRefC - fDewRefC) <> 0.0)
   OR (fTempRefC <> fTempRefC) OR ((fTempRefC - fTempRefC) <> 0.0)
   OR (fTimeRefMin <> fTimeRefMin) OR ((fTimeRefMin - fTimeRefMin) <> 0.0)
   OR (fLimitPct <> fLimitPct) OR ((fLimitPct - fLimitPct) <> 0.0) THEN
    FC_DL_DelubeResidualCarbonCalc := -1.0;  (* 哨兵 -1：输入非有限 / Sentinel -1 non-finite *)
    RETURN;
END_IF
(* 组态域闸：停留时间为除子，三个基准量为比例基，限值须为正 *)
IF (fResidTimeMin <= DL_EPS) OR (fTimeRefMin <= DL_EPS) OR (fLimitPct <= DL_ZERO)
   OR (fLubePct < DL_ZERO) THEN
    FC_DL_DelubeResidualCarbonCalc := -1.0;  (* 哨兵 -1：组态非法 / Sentinel -1 bad config *)
    RETURN;
END_IF
(* 露点修正：露点越高越缺氧，烧除越不完全，残碳升高 *)
fKDew := 1.0 + (fDewPointC - fDewRefC) * DL_DEW_K;
IF fKDew < DL_K_MIN THEN
    fKDew := DL_K_MIN;
ELSIF fKDew > DL_K_MAX THEN
    fKDew := DL_K_MAX;
END_IF
(* 温度修正：温度越低烧除越不完全，残碳升高 *)
fKTmp := 1.0 + (fTempRefC - fZoneTempC) * DL_TMP_K;
IF fKTmp < DL_K_MIN THEN
    fKTmp := DL_K_MIN;
ELSIF fKTmp > DL_K_MAX THEN
    fKTmp := DL_K_MAX;
END_IF
(* 停留时间修正：停留越短烧除越不完全，残碳升高 *)
fKTime := fTimeRefMin / fResidTimeMin;
IF fKTime < DL_K_MIN THEN
    fKTime := DL_K_MIN;
ELSIF fKTime > DL_K_MAX THEN
    fKTime := DL_K_MAX;
END_IF
(* 综合修正系数与残碳估算：分母均已过域闸 *)
fKCoef := fKDew * fKTmp * fKTime;
fResidualPct := fLubePct * fKCoef;
(* 合格判定：残碳不超过限值 *)
xQualified := fResidualPct <= fLimitPct;
xValid := TRUE;                             (* 链路有效 / Chain valid *)
FC_DL_DelubeResidualCarbonCalc := fResidualPct;  (* 返回残碳 [%] / Return residual carbon *)
END_FUNCTION

(* ---- FC_DL_DieCastPorosityRiskIndexCalc.st ---- *)
(*
  Component : FC_DL_DieCastPorosityRiskIndexCalc
  Category  : DL_Device
  Type      : FC
  Complexity: C2
  VERSION   : v1.0.0
  功能      : 压铸气孔风险指数评估：按卷气（压射速度）、模温差、排气能力三因子加权算 0~100 风险指数并给出 1~4 风险等级。
  开源溯源  : 道莅原创 clean-room 自研（无外部代码引用）｜License: MIT
  边界条件  : ① 三个基准量（参考速度、参考温差、参考排气面积）须 > 1e-9，否则返回哨兵 -1；
              ② 各单因子先归一化为 0~100 并双侧钳位，再做加权，避免单因子拉爆总分；
              ③ 排气因子取反向：排气面积越小风险越高。
*)
FUNCTION FC_DL_DieCastPorosityRiskIndexCalc : REAL
VAR_INPUT
    fShotVelMs     : REAL;   (* 空压射速度 [m/s] Dry shot velocity *)
    fVelRefMs      : REAL;   (* 卷气基准速度（工艺窗口上限） [m/s] Velocity reference *)
    fTempDiffK     : REAL;   (* 模面温差 [K] Die surface temperature difference *)
    fTempDiffRefK  : REAL;   (* 温差基准（允许上限） [K] Temperature difference reference *)
    fVentAreaMm2   : REAL;   (* 排气截面积 [mm²] Vent cross-section area *)
    fVentRefMm2    : REAL;   (* 排气基准面积（设计值） [mm²] Vent reference area *)
END_VAR
VAR_OUTPUT
    fRiskIdx    : REAL;   (* 综合气孔风险指数 0~100 [-] Composite porosity risk index *)
    fVelFactor  : REAL;   (* 卷气因子 0~100 [-] Air entrapment factor *)
    fTempFactor : REAL;   (* 温差因子 0~100 [-] Temperature factor *)
    fVentFactor : REAL;   (* 排气因子 0~100 [-] Venting factor *)
    nRiskGrade  : INT;    (* 风险等级 1~4 [-] Risk grade *)
    xValid      : BOOL;   (* 计算有效性标志 [-] Calculation valid flag *)
END_VAR
VAR CONSTANT
    DL_EPS      : REAL := 1.0E-9;   (* 除零判定容差 [无量纲] Divide-by-zero tolerance *)
    DL_PCT_BASE : REAL := 100.0;    (* 百分比基准 [%] Percent base *)
    DL_W_VEL    : REAL := 0.40;     (* 卷气因子权重 [-] Velocity factor weight *)
    DL_W_TEMP   : REAL := 0.35;     (* 温差因子权重 [-] Temperature factor weight *)
    DL_W_VENT   : REAL := 0.25;     (* 排气因子权重 [-] Venting factor weight *)
    DL_ONE      : REAL := 1.0;      (* 单位常数 [-] Unity constant *)
    DL_ZERO     : REAL := 0.0;      (* 零常量 [无量纲] Zero constant *)
END_VAR
VAR
    fRawV : REAL;   (* 卷气因子原始值 [-] Raw velocity factor *)
    fRawT : REAL;   (* 温差因子原始值 [-] Raw temperature factor *)
    fRawE : REAL;   (* 排气因子原始值 [-] Raw venting factor *)
END_VAR
(* 出口预置：六出口统一预置 *)
fRiskIdx := 0.0; fVelFactor := 0.0; fTempFactor := 0.0; fVentFactor := 0.0;
nRiskGrade := 1; xValid := FALSE;
(* 非有限拦截：自反判 NaN，自身差值判 Inf *)
IF (fShotVelMs <> fShotVelMs) OR ((fShotVelMs - fShotVelMs) <> 0.0)
   OR (fTempDiffK <> fTempDiffK) OR ((fTempDiffK - fTempDiffK) <> 0.0)
   OR (fVentAreaMm2 <> fVentAreaMm2) OR ((fVentAreaMm2 - fVentAreaMm2) <> 0.0)
   OR (fVelRefMs <> fVelRefMs) OR ((fVelRefMs - fVelRefMs) <> 0.0)
   OR (fTempDiffRefK <> fTempDiffRefK) OR ((fTempDiffRefK - fTempDiffRefK) <> 0.0)
   OR (fVentRefMm2 <> fVentRefMm2) OR ((fVentRefMm2 - fVentRefMm2) <> 0.0) THEN
    FC_DL_DieCastPorosityRiskIndexCalc := -1.0;  (* 哨兵 -1：输入非有限 / Sentinel -1 non-finite *)
    RETURN;
END_IF
(* 组态域闸：三个基准量全部为除子 *)
IF (fVelRefMs <= DL_EPS) OR (fTempDiffRefK <= DL_EPS) OR (fVentRefMm2 <= DL_EPS)
   OR (fShotVelMs < DL_ZERO) THEN
    FC_DL_DieCastPorosityRiskIndexCalc := -1.0;  (* 哨兵 -1：组态非法 / Sentinel -1 bad config *)
    RETURN;
END_IF
(* 卷气因子：速度越高卷气越重，归一化后双侧钳位 0~100 *)
fRawV := fShotVelMs / fVelRefMs * DL_PCT_BASE;
IF fRawV > DL_PCT_BASE THEN
    fVelFactor := DL_PCT_BASE;
ELSIF fRawV < DL_ZERO THEN
    fVelFactor := DL_ZERO;
ELSE
    fVelFactor := fRawV;
END_IF
(* 温差因子：温差越大热节越重，归一化后双侧钳位 0~100 *)
fRawT := fTempDiffK / fTempDiffRefK * DL_PCT_BASE;
IF fRawT > DL_PCT_BASE THEN
    fTempFactor := DL_PCT_BASE;
ELSIF fRawT < DL_ZERO THEN
    fTempFactor := DL_ZERO;
ELSE
    fTempFactor := fRawT;
END_IF
(* 排气因子：排气面积越小风险越高，取 1 - 面积比 并双侧钳位 *)
fRawE := (DL_ONE - fVentAreaMm2 / fVentRefMm2) * DL_PCT_BASE;
IF fRawE > DL_PCT_BASE THEN
    fVentFactor := DL_PCT_BASE;
ELSIF fRawE < DL_ZERO THEN
    fVentFactor := DL_ZERO;
ELSE
    fVentFactor := fRawE;
END_IF
(* 加权合成：三因子权重之和为 1，结果为 0~100 *)
fRiskIdx := fVelFactor * DL_W_VEL + fTempFactor * DL_W_TEMP + fVentFactor * DL_W_VENT;
(* 风险分级：<25 优 / <50 良 / <75 中 / 其余 差 *)
IF fRiskIdx < 25.0 THEN
    nRiskGrade := 1;
ELSIF fRiskIdx < 50.0 THEN
    nRiskGrade := 2;
ELSIF fRiskIdx < 75.0 THEN
    nRiskGrade := 3;
ELSE
    nRiskGrade := 4;
END_IF
xValid := TRUE;                                  (* 链路有效 / Chain valid *)
FC_DL_DieCastPorosityRiskIndexCalc := fRiskIdx;  (* 返回风险指数 [-] / Return risk index *)
END_FUNCTION

(* ---- FC_DL_DoSalinityPermCalc.st ---- *)
(* ============================================================
   DL_Device / FC_DL_DoSalinityPermCalc ｜ v1.0.0 ｜ 2026-11-25
   功能：溶解氧膜渗透与盐度/温度修正
         C_corr = (C_raw + k_S · S) · K_perm · (1 + k_T · (T − 25)) [mg/L]，
         k_S = 0.084 mg/L 每 ‰（盐度使表观溶解度下降，故加回），k_T = 引脚 %/°C ÷ 100。
   边界：量程上限 ≤ 0 或渗透因子 ≤ 0 → 浓度写 0、返回 FALSE（N1/N3）；
         任一入参非有限 → 浓度写 0、返回 FALSE；盐度 < 0 按 0 处理且 bSalApplied=FALSE；
         C_corr 越出 [0, 上限] → 钳端点并置 bOutOfRange。签名无出口码，闸序即归因序。
         量纲清单（N5）：1 ‰ = 1 g/kg 盐度；k_S = 0.084 mg/L per ‰ = 84 µg/L 每 g/kg；
         回代：S = 35 ‰ 时表观溶解度下降 2.94 mg/L。
   依赖：仅 IEC 61131-3（无外部依赖，纯算术） ｜ 溯源：DLF-D-WATERANA
   验收：C=8.00/T=25/S=0/K=1.0/上限 20/kT=2.0 → 8.00 mg/L、未越限、TRUE；
         S=35 → (8.00 + 2.94) = 10.94 mg/L、bSalApplied=TRUE。
   ============================================================ *)
FUNCTION FC_DL_DoSalinityPermCalc : BOOL
VAR_INPUT
    fDoRaw       : REAL;  // 表读溶解氧浓度 [mg/L] / Dissolved oxygen reading from the probe
    fTempC       : REAL;  // 水温 [°C] / Water temperature in Celsius degrees
    fSalinityPpt : REAL;  // 盐度，有效域 ≥ 0 [‰] / Salinity in parts per thousand
    fPermK       : REAL;  // 膜渗透系标定因子，有效域 > 0 [-] / Membrane permeability calibration factor
    fDoMax       : REAL;  // 量程上限，有效域 > 0 [mg/L] / Upper range limit of the measurement
    fTempCoefPct : REAL;  // 温度修正系数（%/°C，可为负）[%/°C] / Temperature correction coefficient
END_VAR
VAR_OUTPUT
    fDoCorrMgL  : REAL;  // 修正后溶解氧浓度 [mg/L] / Corrected dissolved oxygen concentration
    bOutOfRange : BOOL;  // 修正值被钳到量程端点 [-] / Corrected value clamped to a range end
    bSalApplied : BOOL;  // 盐度修正已生效（盐度 > 0）[-] / Salinity correction actually applied
END_VAR
VAR
    _fSal : REAL;  // 归零后的盐度 [‰] / Normalized salinity
    _fKt  : REAL;  // 温度修正因子 (1 + k_T·(T−25)) [-] / Temperature correction factor
    _fC   : REAL;  // 修正中间值 [mg/L] / Intermediate corrected value
END_VAR
VAR CONSTANT
    DL_DOS_KS   : REAL := 0.084;  // 盐度溶解度系数 [mg/L per ‰] / Salinity solubility coefficient
    DL_DOS_TREF : REAL := 25.0;   // 参考温度 [°C] / Reference temperature
    DL_DOS_HUND : REAL := 100.0;  // 百分比换算系数 [%] / Percent conversion factor
END_VAR

(* 段 0：出口预置安全侧（0 mg/L、两标志置位，N1/N3） *)
FC_DL_DoSalinityPermCalc := FALSE;
fDoCorrMgL := 0.0;  bOutOfRange := TRUE;  bSalApplied := FALSE;

(* 段 1：非有限闸（六个入参全量枚举） *)
IF (fDoRaw <> fDoRaw) OR (fTempC <> fTempC) OR (fSalinityPpt <> fSalinityPpt)
   OR (fPermK <> fPermK) OR (fDoMax <> fDoMax) OR (fTempCoefPct <> fTempCoefPct) THEN RETURN; END_IF

(* 段 2：域闸（量程上限与渗透因子必须为正） *)
IF (fDoMax <= 0.0) OR (fPermK <= 0.0) THEN RETURN; END_IF

(* 段 3：盐度归零（负输入按 0 处理，并如实标记未生效） *)
IF fSalinityPpt > 0.0 THEN
    _fSal := fSalinityPpt;  bSalApplied := TRUE;
ELSE
    _fSal := 0.0;           bSalApplied := FALSE;
END_IF

(* 段 4：温度因子与修正（乘加，除子为常量 100） *)
_fKt := 1.0 + (fTempCoefPct / DL_DOS_HUND) * (fTempC - DL_DOS_TREF);
_fC  := (fDoRaw + DL_DOS_KS * _fSal) * fPermK * _fKt;

(* 段 5：结果复检（非有限保持段 0 安全侧） *)
IF (_fC <> _fC) OR ((_fC - _fC) <> (_fC - _fC)) THEN RETURN; END_IF

(* 段 6：单一出口裁决（判据与出口同源于 _fC，N4/R23） *)
bOutOfRange := ((_fC < 0.0) OR (_fC > fDoMax));
IF _fC < 0.0 THEN
    fDoCorrMgL := 0.0;                  // 负值保护：钳零后上报
ELSIF _fC > fDoMax THEN
    fDoCorrMgL := fDoMax;               // 饱和上报：钳顶后值仍可读
ELSE
    fDoCorrMgL := _fC;
END_IF
FC_DL_DoSalinityPermCalc := TRUE;
END_FUNCTION

(* ---- FC_DL_ElectrostaticVoltageCalc.st ---- *)
(*
  Name: FC_DL_ElectrostaticVoltageCalc
  Category: DL_Device
  Version: 1.0.0
  Round: R89 / 2026-11-25
  开源溯源：clean-room 自研（族 涂装喷涂线，ST 开源生态实测 0 命中，无外部代码引入）
  功能：静电喷涂电压-电流-距离校核：算电场强度（kV/mm），并分别给出电压上限与距离下限判定。
  边界条件：① 四入参全部过非有限闸，任一非有限返回哨兵 -1；
            ② 枪距为电场强度除子，须 50~500 mm，绝无零除；
            ③ 归因分离（R190）：xVoltSafe 只判电压对上限，xDistSafe 只判距离对下限，两判据不合并；
               电场强度仅作诊断输出，超限不并入任一安全位（避免出口归因混淆）；
            ④ 电流 fCurrentUa 仅参与域闸与诊断，不参与安全位（本件不做电流积分判定）。
  量纲自证：kV ÷ mm = kV/mm；电压与上限、距离与下限各自同量纲比较。
*)
FUNCTION FC_DL_ElectrostaticVoltageCalc : REAL
VAR_INPUT
    fDistMm : REAL;         (* 喷枪到工件距离 [mm] Gun-to-part distance [mm] *)
    fVoltKv : REAL;         (* 静电电压 [kV] Electrostatic voltage [kV] *)
    fCurrentUa : REAL;      (* 静电电流 [μA] Electrostatic current [uA] *)
    fVoltMaxKv : REAL;      (* 电压上限 [kV] Voltage ceiling [kV] *)
    fDistMinMm : REAL;      (* 枪距下限 [mm] Distance floor [mm] *)
END_VAR
VAR_OUTPUT
    fFieldKvPerMm : REAL;   (* 电场强度（诊断量） [kV/mm] Field strength [kV/mm] *)
    xVoltSafe : BOOL;       (* 电压不超上限 [-] Voltage within ceiling *)
    xDistSafe : BOOL;       (* 枪距不低于下限 [-] Distance above floor *)
    xValid : BOOL;          (* 计算有效性标志 [-] Calculation valid flag *)
END_VAR
VAR CONSTANT
    DL_EPS : REAL := 1.0E-9;        (* 判据容差 [-] Criterion tolerance *)
    DL_D_MIN : REAL := 50.0;        (* 枪距量程下限 [mm] Distance floor [mm] *)
    DL_D_MAX : REAL := 500.0;       (* 枪距量程上限 [mm] Distance ceiling [mm] *)
    DL_V_MIN : REAL := 1.0;         (* 电压量程下限 [kV] Voltage floor [kV] *)
    DL_V_MAX : REAL := 120.0;       (* 电压量程上限 [kV] Voltage ceiling [kV] *)
    DL_I_MIN : REAL := 0.0;         (* 电流量程下限 [μA] Current floor [uA] *)
    DL_I_MAX : REAL := 200.0;       (* 电流量程上限 [μA] Current ceiling [uA] *)
    DL_VM_MIN : REAL := 1.0;        (* 电压上限下限 [kV] Voltage ceiling floor [kV] *)
    DL_VM_MAX : REAL := 120.0;      (* 电压上限上限 [kV] Voltage ceiling top [kV] *)
    DL_DM_MIN : REAL := 50.0;       (* 枪距下限下限 [mm] Distance floor floor [mm] *)
    DL_DM_MAX : REAL := 500.0;      (* 枪距下限上限 [mm] Distance floor top [mm] *)
END_VAR
(* 出口预置：四出口统一预置（R256） *)
fFieldKvPerMm := 0.0; xVoltSafe := FALSE; xDistSafe := FALSE; xValid := FALSE;
(* 非有限闸：NaN 自反判 + Inf 差值自减判，五入参全枚举（R272） *)
IF (fDistMm <> fDistMm) OR ((fDistMm - fDistMm) <> 0.0)
   OR (fVoltKv <> fVoltKv) OR ((fVoltKv - fVoltKv) <> 0.0)
   OR (fCurrentUa <> fCurrentUa) OR ((fCurrentUa - fCurrentUa) <> 0.0)
   OR (fVoltMaxKv <> fVoltMaxKv) OR ((fVoltMaxKv - fVoltMaxKv) <> 0.0)
   OR (fDistMinMm <> fDistMinMm) OR ((fDistMinMm - fDistMinMm) <> 0.0) THEN
    FC_DL_ElectrostaticVoltageCalc := -1.0; (* 哨兵 -1：入参非有限 / Sentinel -1, non-finite input *)
    RETURN;
END_IF
(* 组态域闸：枪距、电压、电流、两限值逐项定域（枪距为除子） *)
IF (fDistMm < DL_D_MIN) OR (fDistMm > DL_D_MAX)
   OR (fVoltKv < DL_V_MIN) OR (fVoltKv > DL_V_MAX)
   OR (fCurrentUa < DL_I_MIN) OR (fCurrentUa > DL_I_MAX)
   OR (fVoltMaxKv < DL_VM_MIN) OR (fVoltMaxKv > DL_VM_MAX)
   OR (fDistMinMm < DL_DM_MIN) OR (fDistMinMm > DL_DM_MAX) THEN
    FC_DL_ElectrostaticVoltageCalc := -1.0; (* 哨兵 -1：组态非法 / Sentinel -1, bad configuration *)
    RETURN;
END_IF
(* 电场强度：kV ÷ mm = kV/mm，枪距已过下限闸绝无零除 *)
fFieldKvPerMm := fVoltKv / fDistMm;
(* 归因唯一：电压判据只比电压上限；距离判据只比距离下限 *)
xVoltSafe := fVoltKv <= fVoltMaxKv;
xDistSafe := fDistMm >= fDistMinMm;
xValid := TRUE;                             (* 链路有效 / Chain valid *)
FC_DL_ElectrostaticVoltageCalc := fFieldKvPerMm;
END_FUNCTION

(* ---- FC_DL_FiberCoolingAirflowCalc.st ---- *)
// FC_DL_FiberCoolingAirflowCalc v1.0.0
// 开源溯源：clean-room 自研（族 DL_Device，ST 生态实测 0 命中，无外部代码引入）
(*
  功能: 丝束冷却风量：ΔT = 出风 − 进风 [K]，ΔT ≤ 0.5 K 拒收（换热量不可分辨）；
        质量流量 = Q[kW]/(1.005·ΔT) [kg/s]（1.005 为空气定压比热 kJ/(kg·K)），
        体积风量 = 质量流量/密度×3600 [m³/h]。
  邻件/码位: 与 FC_DL_BushingPowerBalanceCalc 同属热平衡链（丝束冷却侧 vs 漏板本体散热）；
             16#0002_9228 = 非有限、热量/密度非正或温差不足 0.5 K 拒收。
*)
FUNCTION FC_DL_FiberCoolingAirflowCalc : REAL
VAR_INPUT
    fHeatToRemove  : REAL := 8.0;       // 需带走热量 [kW]，域 > 0 / Heat to remove [kW]
    fAirInletTemp  : REAL := 30.0;      // 进风温度 [°C] / Inlet air temperature [degC]
    fAirOutletTemp : REAL := 45.0;      // 出风温度 [°C] / Outlet air temperature [degC]
    fAirDensity    : REAL := 1.15;      // 空气密度 [kg/m³]，域 > 0 / Air density [kg/m^3]
END_VAR
VAR_OUTPUT
    fAirflowM3h : REAL;                 // 体积风量 [m³/h] / Volumetric airflow [m^3/h]
    bValid      : BOOL;                 // 结果有效回执 [-] / Result validity receipt
    uErrorId    : UDINT;                // 事件码，0 = 无事件 / Event code
END_VAR
VAR
    fDeltaT : REAL := 0.0;              // 进出风温差 [K] / Temperature rise [K]
END_VAR
// 段 0：全路径出口安全缺省 / Safe defaults on all outlets
fAirflowM3h := 0.0;                 // 风量缺省零 / Airflow default zero
bValid := FALSE;                    // 有效回执预清 / Validity preset clear
uErrorId := 16#0000;                // 事件码预清 / Event code preset clear
FC_DL_FiberCoolingAirflowCalc := 0.0;   // 返回值缺省零（镜像风量）/ Return default zero
// 段 1：非有限闸（四入参全枚举）/ Non-finite gate over all inputs
IF (fHeatToRemove <> fHeatToRemove) OR (fAirInletTemp <> fAirInletTemp)
   OR (fAirOutletTemp <> fAirOutletTemp) OR (fAirDensity <> fAirDensity)
   OR (ABS(fHeatToRemove) >= 3.0E38) OR (ABS(fAirInletTemp) >= 3.0E38)
   OR (ABS(fAirOutletTemp) >= 3.0E38) OR (ABS(fAirDensity) >= 3.0E38) THEN
    uErrorId := 16#0002_9228;   // 入参非有限拒收 / Non-finite input reject
    RETURN;
END_IF
// 段 2：域闸（热量与密度为正 + 温差可分辨，R4）/ Domain gate
IF (fHeatToRemove <= 1.0E-6) OR (fAirDensity <= 1.0E-6) THEN
    uErrorId := 16#0002_9228;   // 热量或密度非正 / Non-positive heat or density
    RETURN;
END_IF
fDeltaT := fAirOutletTemp - fAirInletTemp;                      // 温差 [K] / Temperature rise
IF fDeltaT <= 0.5 THEN
    uErrorId := 16#0002_9228;   // 温差不足 0.5 K，风量解发散 / Rise too small
    RETURN;
END_IF
// 段 3：主计算（质量流量 → 体积风量）/ Main computation
fAirflowM3h := (fHeatToRemove / (1.005 * fDeltaT)) / fAirDensity * 3600.0;  // [m³/h] / Airflow
// 段 4：出口闸（非有限复核 + 正数复核）/ Outlet gate
IF (fAirflowM3h <> fAirflowM3h) OR (ABS(fAirflowM3h) >= 3.0E38) OR (fAirflowM3h <= 0.0) THEN
    fAirflowM3h := 0.0;         // 复核失败回缺省 / Fallback on recheck failure
    uErrorId := 16#0002_9228;   // 出口复核拒收 / Output recheck reject
    RETURN;
END_IF
bValid := TRUE;                 // 有效回执 / Validity receipt
FC_DL_FiberCoolingAirflowCalc := fAirflowM3h;   // 返回值镜像风量 / Return mirrors airflow
END_FUNCTION
